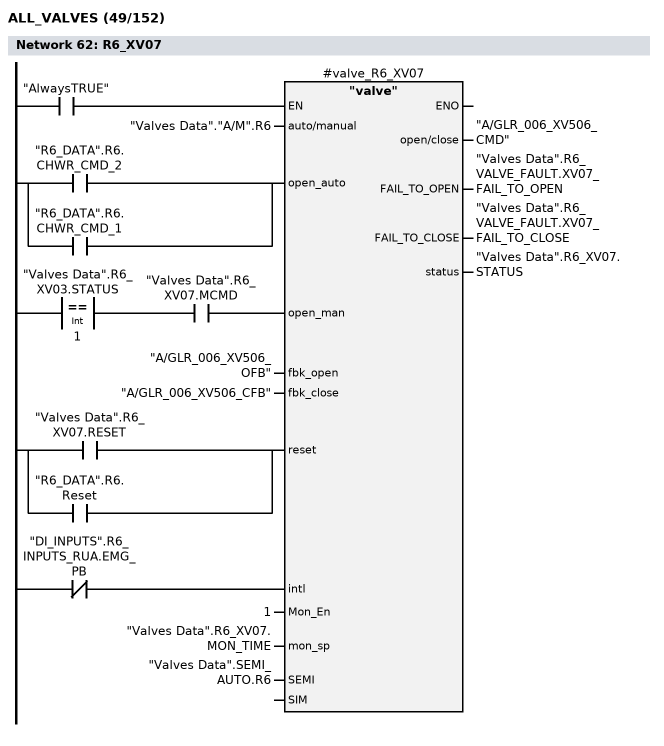
   RUNG wire#powerrail
      Contact( "AlwaysTRUE" )
      #valve_R6_XV07(open_auto := wire#w1, open_man := wire#w2, reset := wire#w3, intl := wire#w4, "auto/manual" := "Valves Data"."A/M".R6, fbk_open := "A/GLR_006_XV506_OFB", fbk_close := "A/GLR_006_XV506_CFB", Mon_En := 1, mon_sp := "Valves Data".R6_XV07.MON_TIME, SEMI := "Valves Data".SEMI_AUTO.R6, SIM :=, "open/close" => "A/GLR_006_XV506_CMD", FAIL_TO_OPEN => "Valves Data".R6_VALVE_FAULT.XV07_FAIL_TO_OPEN, FAIL_TO_CLOSE => "Valves Data".R6_VALVE_FAULT.XV07_FAIL_TO_CLOSE, status => "Valves Data".R6_XV07.STATUS)
   END_RUNG
   RUNG wire#powerrail
      Contact( "R6_DATA".R6.CHWR_CMD_2 )
   END_RUNG wire#w1
   RUNG wire#powerrail
      Contact( "R6_DATA".R6.CHWR_CMD_1 )
   END_RUNG wire#w1
   RUNG wire#powerrail
      { S7_Templates := "SrcType := Int" } EQ_Contact(in1 := "Valves Data".R6_XV03.STATUS, in2 := 1)
      Contact( "Valves Data".R6_XV07.MCMD )
   END_RUNG wire#w2
   RUNG wire#powerrail
      Contact( "Valves Data".R6_XV07.RESET )
   END_RUNG wire#w3
   RUNG wire#powerrail
      Contact( "R6_DATA".R6.Reset )
   END_RUNG wire#w3
   RUNG wire#powerrail
      I_Contact( "DI_INPUTS".R6_INPUTS_RUA.EMG_PB )
   END_RUNG wire#w4
   // the same network as SCL:
   IF "AlwaysTRUE" THEN
       #valve_R6_XV07("auto/manual" := "Valves Data"."A/M".R6,   // "valve"
                      open_auto := "R6_DATA".R6.CHWR_CMD_2 OR "R6_DATA".R6.CHWR_CMD_1,
                      open_man := ("Valves Data".R6_XV03.STATUS = 1) AND "Valves Data".R6_XV07.MCMD,
                      fbk_open := "A/GLR_006_XV506_OFB",
                      fbk_close := "A/GLR_006_XV506_CFB",
                      reset := "Valves Data".R6_XV07.RESET OR "R6_DATA".R6.Reset,
                      intl := NOT "DI_INPUTS".R6_INPUTS_RUA.EMG_PB,
                      Mon_En := 1,
                      mon_sp := "Valves Data".R6_XV07.MON_TIME,
                      SEMI := "Valves Data".SEMI_AUTO.R6,
                      "open/close" => "A/GLR_006_XV506_CMD",
                      FAIL_TO_OPEN => "Valves Data".R6_VALVE_FAULT.XV07_FAIL_TO_OPEN,
                      FAIL_TO_CLOSE => "Valves Data".R6_VALVE_FAULT.XV07_FAIL_TO_CLOSE,
                      status => "Valves Data".R6_XV07.STATUS);
   END_IF;
END_REGION

REGION Network 63: R6_XV08
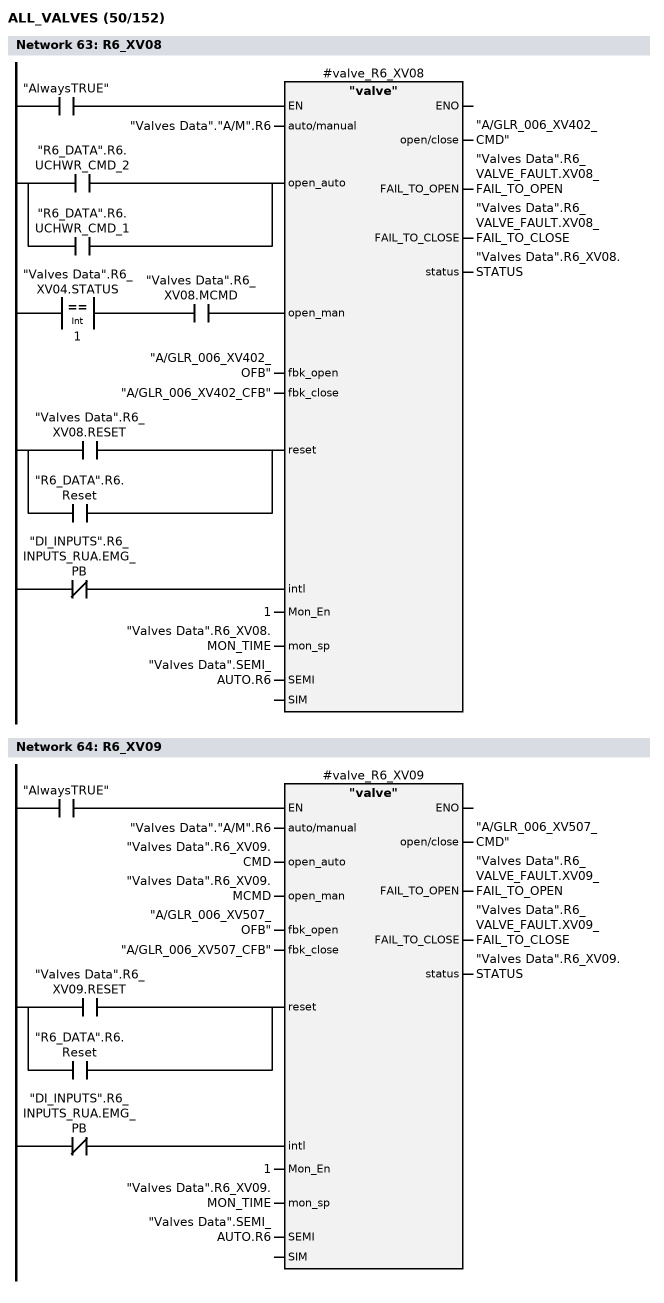
   RUNG wire#powerrail
      Contact( "AlwaysTRUE" )
      #valve_R6_XV08(open_auto := wire#w1, open_man := wire#w2, reset := wire#w3, intl := wire#w4, "auto/manual" := "Valves Data"."A/M".R6, fbk_open := "A/GLR_006_XV402_OFB", fbk_close := "A/GLR_006_XV402_CFB", Mon_En := 1, mon_sp := "Valves Data".R6_XV08.MON_TIME, SEMI := "Valves Data".SEMI_AUTO.R6, SIM :=, "open/close" => "A/GLR_006_XV402_CMD", FAIL_TO_OPEN => "Valves Data".R6_VALVE_FAULT.XV08_FAIL_TO_OPEN, FAIL_TO_CLOSE => "Valves Data".R6_VALVE_FAULT.XV08_FAIL_TO_CLOSE, status => "Valves Data".R6_XV08.STATUS)
   END_RUNG
   RUNG wire#powerrail
      Contact( "R6_DATA".R6.UCHWR_CMD_2 )
   END_RUNG wire#w1
   RUNG wire#powerrail
      Contact( "R6_DATA".R6.UCHWR_CMD_1 )
   END_RUNG wire#w1
   RUNG wire#powerrail
      { S7_Templates := "SrcType := Int" } EQ_Contact(in1 := "Valves Data".R6_XV04.STATUS, in2 := 1)
      Contact( "Valves Data".R6_XV08.MCMD )
   END_RUNG wire#w2
   RUNG wire#powerrail
      Contact( "Valves Data".R6_XV08.RESET )
   END_RUNG wire#w3
   RUNG wire#powerrail
      Contact( "R6_DATA".R6.Reset )
   END_RUNG wire#w3
   RUNG wire#powerrail
      I_Contact( "DI_INPUTS".R6_INPUTS_RUA.EMG_PB )
   END_RUNG wire#w4
   // the same network as SCL:
   IF "AlwaysTRUE" THEN
       #valve_R6_XV08("auto/manual" := "Valves Data"."A/M".R6,   // "valve"
                      open_auto := "R6_DATA".R6.UCHWR_CMD_2 OR "R6_DATA".R6.UCHWR_CMD_1,
                      open_man := ("Valves Data".R6_XV04.STATUS = 1) AND "Valves Data".R6_XV08.MCMD,
                      fbk_open := "A/GLR_006_XV402_OFB",
                      fbk_close := "A/GLR_006_XV402_CFB",
                      reset := "Valves Data".R6_XV08.RESET OR "R6_DATA".R6.Reset,
                      intl := NOT "DI_INPUTS".R6_INPUTS_RUA.EMG_PB,
                      Mon_En := 1,
                      mon_sp := "Valves Data".R6_XV08.MON_TIME,
                      SEMI := "Valves Data".SEMI_AUTO.R6,
                      "open/close" => "A/GLR_006_XV402_CMD",
                      FAIL_TO_OPEN => "Valves Data".R6_VALVE_FAULT.XV08_FAIL_TO_OPEN,
                      FAIL_TO_CLOSE => "Valves Data".R6_VALVE_FAULT.XV08_FAIL_TO_CLOSE,
                      status => "Valves Data".R6_XV08.STATUS);
   END_IF;
END_REGION

REGION Network 64: R6_XV09
   RUNG wire#powerrail
      Contact( "AlwaysTRUE" )
      #valve_R6_XV09(reset := wire#w1, intl := wire#w2, "auto/manual" := "Valves Data"."A/M".R6, open_auto := "Valves Data".R6_XV09.CMD, open_man := "Valves Data".R6_XV09.MCMD, fbk_open := "A/GLR_006_XV507_OFB", fbk_close := "A/GLR_006_XV507_CFB", Mon_En := 1, mon_sp := "Valves Data".R6_XV09.MON_TIME, SEMI := "Valves Data".SEMI_AUTO.R6, SIM :=, "open/close" => "A/GLR_006_XV507_CMD", FAIL_TO_OPEN => "Valves Data".R6_VALVE_FAULT.XV09_FAIL_TO_OPEN, FAIL_TO_CLOSE => "Valves Data".R6_VALVE_FAULT.XV09_FAIL_TO_CLOSE, status => "Valves Data".R6_XV09.STATUS)
   END_RUNG
   RUNG wire#powerrail
      Contact( "Valves Data".R6_XV09.RESET )
   END_RUNG wire#w1
   RUNG wire#powerrail
      Contact( "R6_DATA".R6.Reset )
   END_RUNG wire#w1
   RUNG wire#powerrail
      I_Contact( "DI_INPUTS".R6_INPUTS_RUA.EMG_PB )
   END_RUNG wire#w2
   // the same network as SCL:
   IF "AlwaysTRUE" THEN
       #valve_R6_XV09("auto/manual" := "Valves Data"."A/M".R6,   // "valve"
                      open_auto := "Valves Data".R6_XV09.CMD,
                      open_man := "Valves Data".R6_XV09.MCMD,
                      fbk_open := "A/GLR_006_XV507_OFB",
                      fbk_close := "A/GLR_006_XV507_CFB",
                      reset := "Valves Data".R6_XV09.RESET OR "R6_DATA".R6.Reset,
                      intl := NOT "DI_INPUTS".R6_INPUTS_RUA.EMG_PB,
                      Mon_En := 1,
                      mon_sp := "Valves Data".R6_XV09.MON_TIME,
                      SEMI := "Valves Data".SEMI_AUTO.R6,
                      "open/close" => "A/GLR_006_XV507_CMD",
                      FAIL_TO_OPEN => "Valves Data".R6_VALVE_FAULT.XV09_FAIL_TO_OPEN,
                      FAIL_TO_CLOSE => "Valves Data".R6_VALVE_FAULT.XV09_FAIL_TO_CLOSE,
                      status => "Valves Data".R6_XV09.STATUS);
   END_IF;
END_REGION

REGION Network 65: R6_XV10
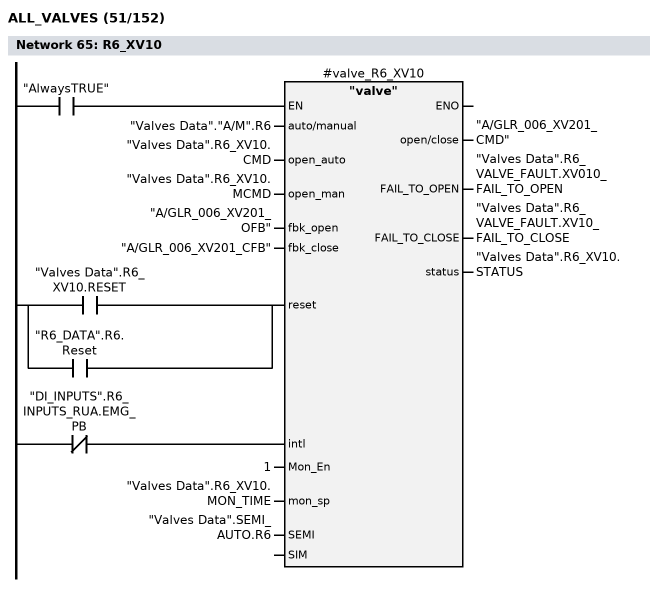
   RUNG wire#powerrail
      Contact( "AlwaysTRUE" )
      #valve_R6_XV10(reset := wire#w1, intl := wire#w2, "auto/manual" := "Valves Data"."A/M".R6, open_auto := "Valves Data".R6_XV10.CMD, open_man := "Valves Data".R6_XV10.MCMD, fbk_open := "A/GLR_006_XV201_OFB", fbk_close := "A/GLR_006_XV201_CFB", Mon_En := 1, mon_sp := "Valves Data".R6_XV10.MON_TIME, SEMI := "Valves Data".SEMI_AUTO.R6, SIM :=, "open/close" => "A/GLR_006_XV201_CMD", FAIL_TO_OPEN => "Valves Data".R6_VALVE_FAULT.XV010_FAIL_TO_OPEN, FAIL_TO_CLOSE => "Valves Data".R6_VALVE_FAULT.XV10_FAIL_TO_CLOSE, status => "Valves Data".R6_XV10.STATUS)
   END_RUNG
   RUNG wire#powerrail
      Contact( "Valves Data".R6_XV10.RESET )
   END_RUNG wire#w1
   RUNG wire#powerrail
      Contact( "R6_DATA".R6.Reset )
   END_RUNG wire#w1
   RUNG wire#powerrail
      I_Contact( "DI_INPUTS".R6_INPUTS_RUA.EMG_PB )
   END_RUNG wire#w2
   // the same network as SCL:
   IF "AlwaysTRUE" THEN
       #valve_R6_XV10("auto/manual" := "Valves Data"."A/M".R6,   // "valve"
                      open_auto := "Valves Data".R6_XV10.CMD,
                      open_man := "Valves Data".R6_XV10.MCMD,
                      fbk_open := "A/GLR_006_XV201_OFB",
                      fbk_close := "A/GLR_006_XV201_CFB",
                      reset := "Valves Data".R6_XV10.RESET OR "R6_DATA".R6.Reset,
                      intl := NOT "DI_INPUTS".R6_INPUTS_RUA.EMG_PB,
                      Mon_En := 1,
                      mon_sp := "Valves Data".R6_XV10.MON_TIME,
                      SEMI := "Valves Data".SEMI_AUTO.R6,
                      "open/close" => "A/GLR_006_XV201_CMD",
                      FAIL_TO_OPEN => "Valves Data".R6_VALVE_FAULT.XV010_FAIL_TO_OPEN,
                      FAIL_TO_CLOSE => "Valves Data".R6_VALVE_FAULT.XV10_FAIL_TO_CLOSE,
                      status => "Valves Data".R6_XV10.STATUS);
   END_IF;
END_REGION

REGION Network 66: ****REACTOR_07****
END_REGION

REGION Network 67: R7_XV01
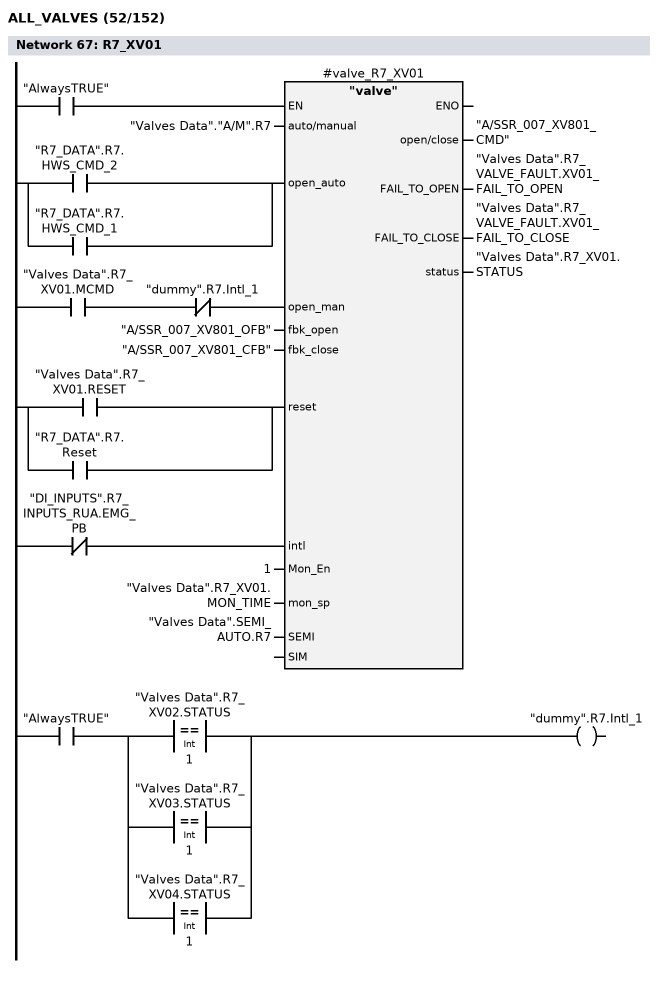
   RUNG wire#powerrail
      Contact( "AlwaysTRUE" )
      #valve_R7_XV01(open_auto := wire#w1, open_man := wire#w2, reset := wire#w3, intl := wire#w4, "auto/manual" := "Valves Data"."A/M".R7, fbk_open := "A/SSR_007_XV801_OFB", fbk_close := "A/SSR_007_XV801_CFB", Mon_En := 1, mon_sp := "Valves Data".R7_XV01.MON_TIME, SEMI := "Valves Data".SEMI_AUTO.R7, SIM :=, "open/close" => "A/SSR_007_XV801_CMD", FAIL_TO_OPEN => "Valves Data".R7_VALVE_FAULT.XV01_FAIL_TO_OPEN, FAIL_TO_CLOSE => "Valves Data".R7_VALVE_FAULT.XV01_FAIL_TO_CLOSE, status => "Valves Data".R7_XV01.STATUS)
   END_RUNG
   RUNG wire#powerrail
      Contact( "R7_DATA".R7.HWS_CMD_2 )
   END_RUNG wire#w1
   RUNG wire#powerrail
      Contact( "R7_DATA".R7.HWS_CMD_1 )
   END_RUNG wire#w1
   RUNG wire#powerrail
      Contact( "Valves Data".R7_XV01.MCMD )
      I_Contact( "dummy".R7.Intl_1 )
   END_RUNG wire#w2
   RUNG wire#powerrail
      Contact( "Valves Data".R7_XV01.RESET )
   END_RUNG wire#w3
   RUNG wire#powerrail
      Contact( "R7_DATA".R7.Reset )
   END_RUNG wire#w3
   RUNG wire#powerrail
      I_Contact( "DI_INPUTS".R7_INPUTS_RUA.EMG_PB )
   END_RUNG wire#w4
   RUNG wire#powerrail
      Contact( "AlwaysTRUE" )
      wire#w5
      { S7_Templates := "SrcType := Int" } EQ_Contact(in1 := "Valves Data".R7_XV02.STATUS, in2 := 1)
      wire#w6
      Coil( "dummy".R7.Intl_1 )
   END_RUNG
   RUNG wire#w5
      { S7_Templates := "SrcType := Int" } EQ_Contact(in1 := "Valves Data".R7_XV03.STATUS, in2 := 1)
   END_RUNG wire#w6
   RUNG wire#w5
      { S7_Templates := "SrcType := Int" } EQ_Contact(in1 := "Valves Data".R7_XV04.STATUS, in2 := 1)
   END_RUNG wire#w6
   // the same network as SCL:
   IF "AlwaysTRUE" THEN
       #valve_R7_XV01("auto/manual" := "Valves Data"."A/M".R7,   // "valve"
                      open_auto := "R7_DATA".R7.HWS_CMD_2 OR "R7_DATA".R7.HWS_CMD_1,
                      open_man := "Valves Data".R7_XV01.MCMD AND NOT "dummy".R7.Intl_1,
                      fbk_open := "A/SSR_007_XV801_OFB",
                      fbk_close := "A/SSR_007_XV801_CFB",
                      reset := "Valves Data".R7_XV01.RESET OR "R7_DATA".R7.Reset,
                      intl := NOT "DI_INPUTS".R7_INPUTS_RUA.EMG_PB,
                      Mon_En := 1,
                      mon_sp := "Valves Data".R7_XV01.MON_TIME,
                      SEMI := "Valves Data".SEMI_AUTO.R7,
                      "open/close" => "A/SSR_007_XV801_CMD",
                      FAIL_TO_OPEN => "Valves Data".R7_VALVE_FAULT.XV01_FAIL_TO_OPEN,
                      FAIL_TO_CLOSE => "Valves Data".R7_VALVE_FAULT.XV01_FAIL_TO_CLOSE,
                      status => "Valves Data".R7_XV01.STATUS);
   END_IF;
   "dummy".R7.Intl_1 := "AlwaysTRUE" AND (("Valves Data".R7_XV02.STATUS = 1) OR ("Valves Data".R7_XV03.STATUS = 1) OR ("Valves Data".R7_XV04.STATUS = 1));
END_REGION

REGION Network 68: R7_XV02
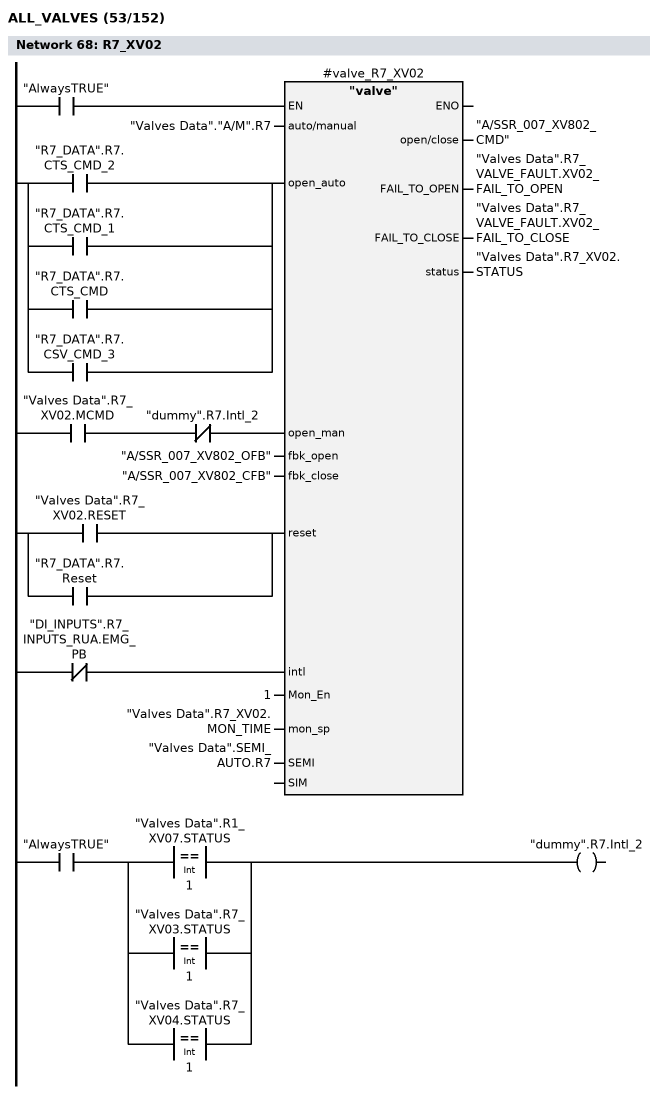
   RUNG wire#powerrail
      Contact( "AlwaysTRUE" )
      #valve_R7_XV02(open_auto := wire#w1, open_man := wire#w2, reset := wire#w3, intl := wire#w4, "auto/manual" := "Valves Data"."A/M".R7, fbk_open := "A/SSR_007_XV802_OFB", fbk_close := "A/SSR_007_XV802_CFB", Mon_En := 1, mon_sp := "Valves Data".R7_XV02.MON_TIME, SEMI := "Valves Data".SEMI_AUTO.R7, SIM :=, "open/close" => "A/SSR_007_XV802_CMD", FAIL_TO_OPEN => "Valves Data".R7_VALVE_FAULT.XV02_FAIL_TO_OPEN, FAIL_TO_CLOSE => "Valves Data".R7_VALVE_FAULT.XV02_FAIL_TO_CLOSE, status => "Valves Data".R7_XV02.STATUS)
   END_RUNG
   RUNG wire#powerrail
      Contact( "R7_DATA".R7.CTS_CMD_2 )
   END_RUNG wire#w1
   RUNG wire#powerrail
      Contact( "R7_DATA".R7.CTS_CMD_1 )
   END_RUNG wire#w1
   RUNG wire#powerrail
      Contact( "R7_DATA".R7.CTS_CMD )
   END_RUNG wire#w1
   RUNG wire#powerrail
      Contact( "R7_DATA".R7.CSV_CMD_3 )
   END_RUNG wire#w1
   RUNG wire#powerrail
      Contact( "Valves Data".R7_XV02.MCMD )
      I_Contact( "dummy".R7.Intl_2 )
   END_RUNG wire#w2
   RUNG wire#powerrail
      Contact( "Valves Data".R7_XV02.RESET )
   END_RUNG wire#w3
   RUNG wire#powerrail
      Contact( "R7_DATA".R7.Reset )
   END_RUNG wire#w3
   RUNG wire#powerrail
      I_Contact( "DI_INPUTS".R7_INPUTS_RUA.EMG_PB )
   END_RUNG wire#w4
   RUNG wire#powerrail
      Contact( "AlwaysTRUE" )
      wire#w5
      { S7_Templates := "SrcType := Int" } EQ_Contact(in1 := "Valves Data".R1_XV07.STATUS, in2 := 1)
      wire#w6
      Coil( "dummy".R7.Intl_2 )
   END_RUNG
   RUNG wire#w5
      { S7_Templates := "SrcType := Int" } EQ_Contact(in1 := "Valves Data".R7_XV03.STATUS, in2 := 1)
   END_RUNG wire#w6
   RUNG wire#w5
      { S7_Templates := "SrcType := Int" } EQ_Contact(in1 := "Valves Data".R7_XV04.STATUS, in2 := 1)
   END_RUNG wire#w6
   // the same network as SCL:
   IF "AlwaysTRUE" THEN
       #valve_R7_XV02("auto/manual" := "Valves Data"."A/M".R7,   // "valve"
                      open_auto := "R7_DATA".R7.CTS_CMD_2 OR "R7_DATA".R7.CTS_CMD_1 OR "R7_DATA".R7.CTS_CMD OR "R7_DATA".R7.CSV_CMD_3,
                      open_man := "Valves Data".R7_XV02.MCMD AND NOT "dummy".R7.Intl_2,
                      fbk_open := "A/SSR_007_XV802_OFB",
                      fbk_close := "A/SSR_007_XV802_CFB",
                      reset := "Valves Data".R7_XV02.RESET OR "R7_DATA".R7.Reset,
                      intl := NOT "DI_INPUTS".R7_INPUTS_RUA.EMG_PB,
                      Mon_En := 1,
                      mon_sp := "Valves Data".R7_XV02.MON_TIME,
                      SEMI := "Valves Data".SEMI_AUTO.R7,
                      "open/close" => "A/SSR_007_XV802_CMD",
                      FAIL_TO_OPEN => "Valves Data".R7_VALVE_FAULT.XV02_FAIL_TO_OPEN,
                      FAIL_TO_CLOSE => "Valves Data".R7_VALVE_FAULT.XV02_FAIL_TO_CLOSE,
                      status => "Valves Data".R7_XV02.STATUS);
   END_IF;
   "dummy".R7.Intl_2 := "AlwaysTRUE" AND (("Valves Data".R1_XV07.STATUS = 1) OR ("Valves Data".R7_XV03.STATUS = 1) OR ("Valves Data".R7_XV04.STATUS = 1));
END_REGION

REGION Network 69: R7_XV03
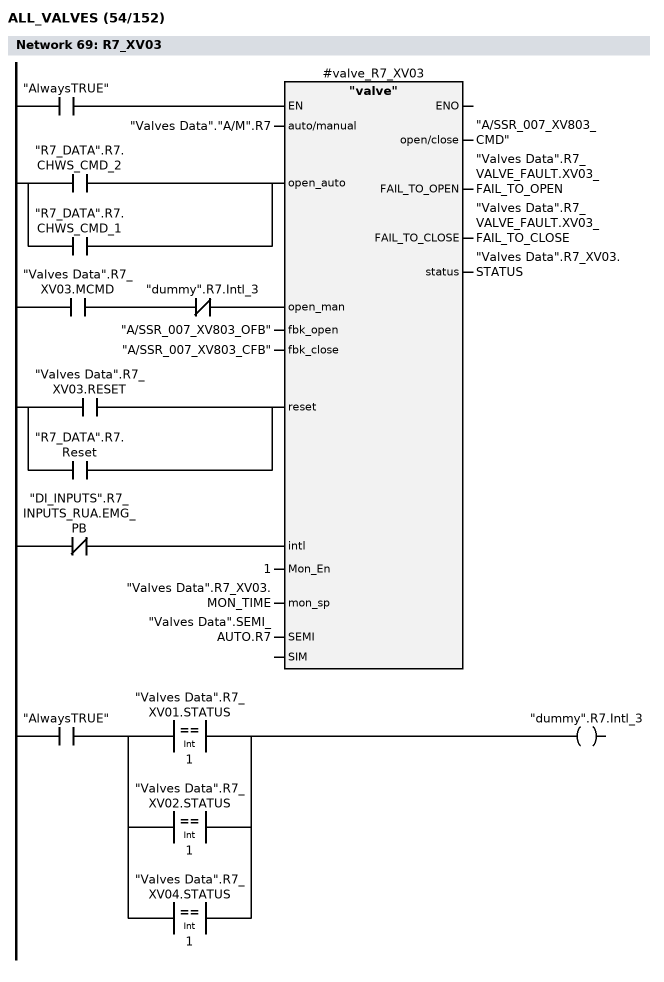
   RUNG wire#powerrail
      Contact( "AlwaysTRUE" )
      #valve_R7_XV03(open_auto := wire#w1, open_man := wire#w2, reset := wire#w3, intl := wire#w4, "auto/manual" := "Valves Data"."A/M".R7, fbk_open := "A/SSR_007_XV803_OFB", fbk_close := "A/SSR_007_XV803_CFB", Mon_En := 1, mon_sp := "Valves Data".R7_XV03.MON_TIME, SEMI := "Valves Data".SEMI_AUTO.R7, SIM :=, "open/close" => "A/SSR_007_XV803_CMD", FAIL_TO_OPEN => "Valves Data".R7_VALVE_FAULT.XV03_FAIL_TO_OPEN, FAIL_TO_CLOSE => "Valves Data".R7_VALVE_FAULT.XV03_FAIL_TO_CLOSE, status => "Valves Data".R7_XV03.STATUS)
   END_RUNG
   RUNG wire#powerrail
      Contact( "R7_DATA".R7.CHWS_CMD_2 )
   END_RUNG wire#w1
   RUNG wire#powerrail
      Contact( "R7_DATA".R7.CHWS_CMD_1 )
   END_RUNG wire#w1
   RUNG wire#powerrail
      Contact( "Valves Data".R7_XV03.MCMD )
      I_Contact( "dummy".R7.Intl_3 )
   END_RUNG wire#w2
   RUNG wire#powerrail
      Contact( "Valves Data".R7_XV03.RESET )
   END_RUNG wire#w3
   RUNG wire#powerrail
      Contact( "R7_DATA".R7.Reset )
   END_RUNG wire#w3
   RUNG wire#powerrail
      I_Contact( "DI_INPUTS".R7_INPUTS_RUA.EMG_PB )
   END_RUNG wire#w4
   RUNG wire#powerrail
      Contact( "AlwaysTRUE" )
      wire#w5
      { S7_Templates := "SrcType := Int" } EQ_Contact(in1 := "Valves Data".R7_XV01.STATUS, in2 := 1)
      wire#w6
      Coil( "dummy".R7.Intl_3 )
   END_RUNG
   RUNG wire#w5
      { S7_Templates := "SrcType := Int" } EQ_Contact(in1 := "Valves Data".R7_XV02.STATUS, in2 := 1)
   END_RUNG wire#w6
   RUNG wire#w5
      { S7_Templates := "SrcType := Int" } EQ_Contact(in1 := "Valves Data".R7_XV04.STATUS, in2 := 1)
   END_RUNG wire#w6
   // the same network as SCL:
   IF "AlwaysTRUE" THEN
       #valve_R7_XV03("auto/manual" := "Valves Data"."A/M".R7,   // "valve"
                      open_auto := "R7_DATA".R7.CHWS_CMD_2 OR "R7_DATA".R7.CHWS_CMD_1,
                      open_man := "Valves Data".R7_XV03.MCMD AND NOT "dummy".R7.Intl_3,
                      fbk_open := "A/SSR_007_XV803_OFB",
                      fbk_close := "A/SSR_007_XV803_CFB",
                      reset := "Valves Data".R7_XV03.RESET OR "R7_DATA".R7.Reset,
                      intl := NOT "DI_INPUTS".R7_INPUTS_RUA.EMG_PB,
                      Mon_En := 1,
                      mon_sp := "Valves Data".R7_XV03.MON_TIME,
                      SEMI := "Valves Data".SEMI_AUTO.R7,
                      "open/close" => "A/SSR_007_XV803_CMD",
                      FAIL_TO_OPEN => "Valves Data".R7_VALVE_FAULT.XV03_FAIL_TO_OPEN,
                      FAIL_TO_CLOSE => "Valves Data".R7_VALVE_FAULT.XV03_FAIL_TO_CLOSE,
                      status => "Valves Data".R7_XV03.STATUS);
   END_IF;
   "dummy".R7.Intl_3 := "AlwaysTRUE" AND (("Valves Data".R7_XV01.STATUS = 1) OR ("Valves Data".R7_XV02.STATUS = 1) OR ("Valves Data".R7_XV04.STATUS = 1));
END_REGION

REGION Network 70: R7_XV04
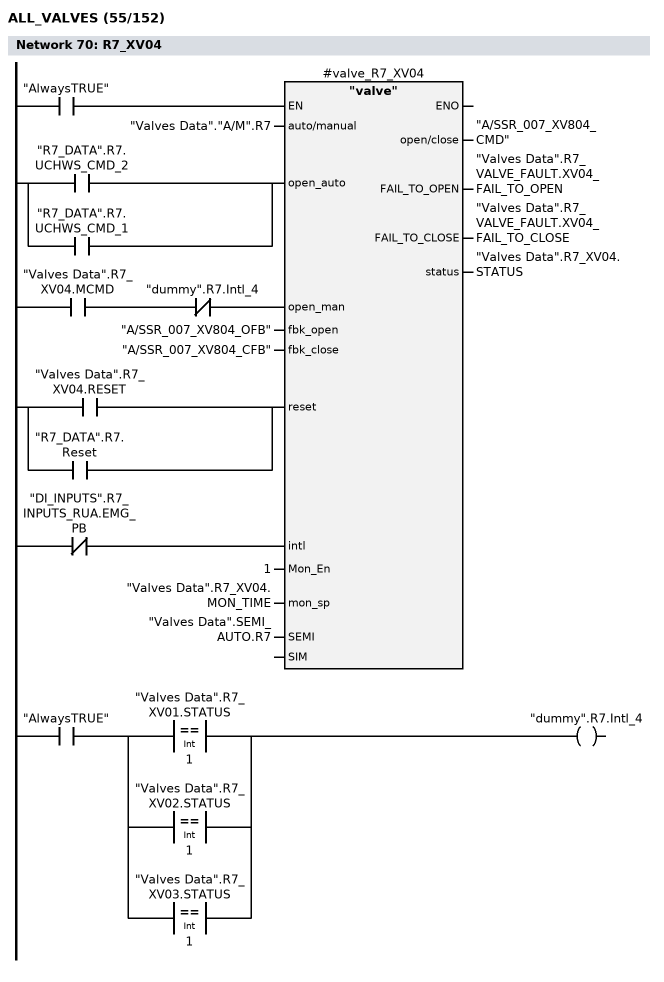
   RUNG wire#powerrail
      Contact( "AlwaysTRUE" )
      #valve_R7_XV04(open_auto := wire#w1, open_man := wire#w2, reset := wire#w3, intl := wire#w4, "auto/manual" := "Valves Data"."A/M".R7, fbk_open := "A/SSR_007_XV804_OFB", fbk_close := "A/SSR_007_XV804_CFB", Mon_En := 1, mon_sp := "Valves Data".R7_XV04.MON_TIME, SEMI := "Valves Data".SEMI_AUTO.R7, SIM :=, "open/close" => "A/SSR_007_XV804_CMD", FAIL_TO_OPEN => "Valves Data".R7_VALVE_FAULT.XV04_FAIL_TO_OPEN, FAIL_TO_CLOSE => "Valves Data".R7_VALVE_FAULT.XV04_FAIL_TO_CLOSE, status => "Valves Data".R7_XV04.STATUS)
   END_RUNG
   RUNG wire#powerrail
      Contact( "R7_DATA".R7.UCHWS_CMD_2 )
   END_RUNG wire#w1
   RUNG wire#powerrail
      Contact( "R7_DATA".R7.UCHWS_CMD_1 )
   END_RUNG wire#w1
   RUNG wire#powerrail
      Contact( "Valves Data".R7_XV04.MCMD )
      I_Contact( "dummy".R7.Intl_4 )
   END_RUNG wire#w2
   RUNG wire#powerrail
      Contact( "Valves Data".R7_XV04.RESET )
   END_RUNG wire#w3
   RUNG wire#powerrail
      Contact( "R7_DATA".R7.Reset )
   END_RUNG wire#w3
   RUNG wire#powerrail
      I_Contact( "DI_INPUTS".R7_INPUTS_RUA.EMG_PB )
   END_RUNG wire#w4
   RUNG wire#powerrail
      Contact( "AlwaysTRUE" )
      wire#w5
      { S7_Templates := "SrcType := Int" } EQ_Contact(in1 := "Valves Data".R7_XV01.STATUS, in2 := 1)
      wire#w6
      Coil( "dummy".R7.Intl_4 )
   END_RUNG
   RUNG wire#w5
      { S7_Templates := "SrcType := Int" } EQ_Contact(in1 := "Valves Data".R7_XV02.STATUS, in2 := 1)
   END_RUNG wire#w6
   RUNG wire#w5
      { S7_Templates := "SrcType := Int" } EQ_Contact(in1 := "Valves Data".R7_XV03.STATUS, in2 := 1)
   END_RUNG wire#w6
   // the same network as SCL:
   IF "AlwaysTRUE" THEN
       #valve_R7_XV04("auto/manual" := "Valves Data"."A/M".R7,   // "valve"
                      open_auto := "R7_DATA".R7.UCHWS_CMD_2 OR "R7_DATA".R7.UCHWS_CMD_1,
                      open_man := "Valves Data".R7_XV04.MCMD AND NOT "dummy".R7.Intl_4,
                      fbk_open := "A/SSR_007_XV804_OFB",
                      fbk_close := "A/SSR_007_XV804_CFB",
                      reset := "Valves Data".R7_XV04.RESET OR "R7_DATA".R7.Reset,
                      intl := NOT "DI_INPUTS".R7_INPUTS_RUA.EMG_PB,
                      Mon_En := 1,
                      mon_sp := "Valves Data".R7_XV04.MON_TIME,
                      SEMI := "Valves Data".SEMI_AUTO.R7,
                      "open/close" => "A/SSR_007_XV804_CMD",
                      FAIL_TO_OPEN => "Valves Data".R7_VALVE_FAULT.XV04_FAIL_TO_OPEN,
                      FAIL_TO_CLOSE => "Valves Data".R7_VALVE_FAULT.XV04_FAIL_TO_CLOSE,
                      status => "Valves Data".R7_XV04.STATUS);
   END_IF;
   "dummy".R7.Intl_4 := "AlwaysTRUE" AND (("Valves Data".R7_XV01.STATUS = 1) OR ("Valves Data".R7_XV02.STATUS = 1) OR ("Valves Data".R7_XV03.STATUS = 1));
END_REGION

REGION Network 71: R7_XV05
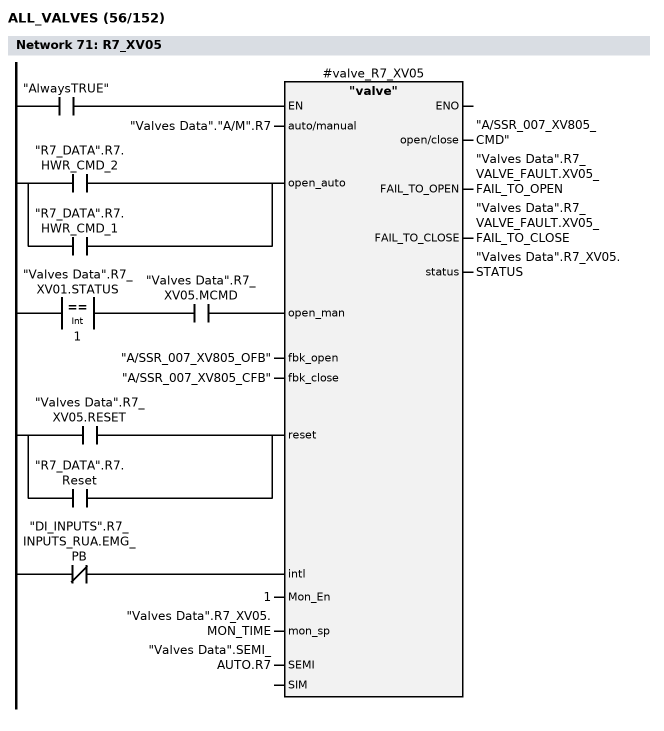
   RUNG wire#powerrail
      Contact( "AlwaysTRUE" )
      #valve_R7_XV05(open_auto := wire#w1, open_man := wire#w2, reset := wire#w3, intl := wire#w4, "auto/manual" := "Valves Data"."A/M".R7, fbk_open := "A/SSR_007_XV805_OFB", fbk_close := "A/SSR_007_XV805_CFB", Mon_En := 1, mon_sp := "Valves Data".R7_XV05.MON_TIME, SEMI := "Valves Data".SEMI_AUTO.R7, SIM :=, "open/close" => "A/SSR_007_XV805_CMD", FAIL_TO_OPEN => "Valves Data".R7_VALVE_FAULT.XV05_FAIL_TO_OPEN, FAIL_TO_CLOSE => "Valves Data".R7_VALVE_FAULT.XV05_FAIL_TO_CLOSE, status => "Valves Data".R7_XV05.STATUS)
   END_RUNG
   RUNG wire#powerrail
      Contact( "R7_DATA".R7.HWR_CMD_2 )
   END_RUNG wire#w1
   RUNG wire#powerrail
      Contact( "R7_DATA".R7.HWR_CMD_1 )
   END_RUNG wire#w1
   RUNG wire#powerrail
      { S7_Templates := "SrcType := Int" } EQ_Contact(in1 := "Valves Data".R7_XV01.STATUS, in2 := 1)
      Contact( "Valves Data".R7_XV05.MCMD )
   END_RUNG wire#w2
   RUNG wire#powerrail
      Contact( "Valves Data".R7_XV05.RESET )
   END_RUNG wire#w3
   RUNG wire#powerrail
      Contact( "R7_DATA".R7.Reset )
   END_RUNG wire#w3
   RUNG wire#powerrail
      I_Contact( "DI_INPUTS".R7_INPUTS_RUA.EMG_PB )
   END_RUNG wire#w4
   // the same network as SCL:
   IF "AlwaysTRUE" THEN
       #valve_R7_XV05("auto/manual" := "Valves Data"."A/M".R7,   // "valve"
                      open_auto := "R7_DATA".R7.HWR_CMD_2 OR "R7_DATA".R7.HWR_CMD_1,
                      open_man := ("Valves Data".R7_XV01.STATUS = 1) AND "Valves Data".R7_XV05.MCMD,
                      fbk_open := "A/SSR_007_XV805_OFB",
                      fbk_close := "A/SSR_007_XV805_CFB",
                      reset := "Valves Data".R7_XV05.RESET OR "R7_DATA".R7.Reset,
                      intl := NOT "DI_INPUTS".R7_INPUTS_RUA.EMG_PB,
                      Mon_En := 1,
                      mon_sp := "Valves Data".R7_XV05.MON_TIME,
                      SEMI := "Valves Data".SEMI_AUTO.R7,
                      "open/close" => "A/SSR_007_XV805_CMD",
                      FAIL_TO_OPEN => "Valves Data".R7_VALVE_FAULT.XV05_FAIL_TO_OPEN,
                      FAIL_TO_CLOSE => "Valves Data".R7_VALVE_FAULT.XV05_FAIL_TO_CLOSE,
                      status => "Valves Data".R7_XV05.STATUS);
   END_IF;
END_REGION

REGION Network 72: R7_XV06
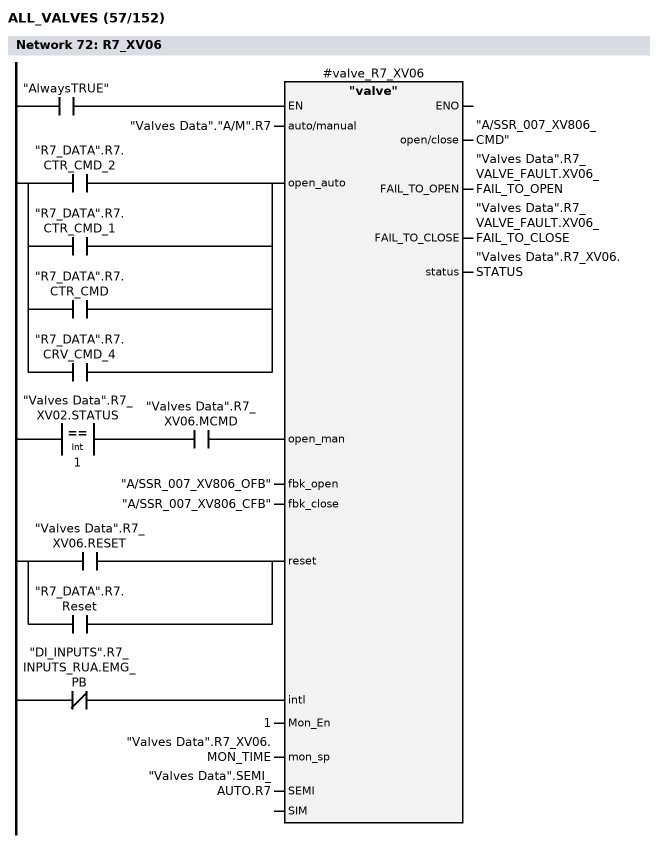
   RUNG wire#powerrail
      Contact( "AlwaysTRUE" )
      #valve_R7_XV06(open_auto := wire#w1, open_man := wire#w2, reset := wire#w3, intl := wire#w4, "auto/manual" := "Valves Data"."A/M".R7, fbk_open := "A/SSR_007_XV806_OFB", fbk_close := "A/SSR_007_XV806_CFB", Mon_En := 1, mon_sp := "Valves Data".R7_XV06.MON_TIME, SEMI := "Valves Data".SEMI_AUTO.R7, SIM :=, "open/close" => "A/SSR_007_XV806_CMD", FAIL_TO_OPEN => "Valves Data".R7_VALVE_FAULT.XV06_FAIL_TO_OPEN, FAIL_TO_CLOSE => "Valves Data".R7_VALVE_FAULT.XV06_FAIL_TO_CLOSE, status => "Valves Data".R7_XV06.STATUS)
   END_RUNG
   RUNG wire#powerrail
      Contact( "R7_DATA".R7.CTR_CMD_2 )
   END_RUNG wire#w1
   RUNG wire#powerrail
      Contact( "R7_DATA".R7.CTR_CMD_1 )
   END_RUNG wire#w1
   RUNG wire#powerrail
      Contact( "R7_DATA".R7.CTR_CMD )
   END_RUNG wire#w1
   RUNG wire#powerrail
      Contact( "R7_DATA".R7.CRV_CMD_4 )
   END_RUNG wire#w1
   RUNG wire#powerrail
      { S7_Templates := "SrcType := Int" } EQ_Contact(in1 := "Valves Data".R7_XV02.STATUS, in2 := 1)
      Contact( "Valves Data".R7_XV06.MCMD )
   END_RUNG wire#w2
   RUNG wire#powerrail
      Contact( "Valves Data".R7_XV06.RESET )
   END_RUNG wire#w3
   RUNG wire#powerrail
      Contact( "R7_DATA".R7.Reset )
   END_RUNG wire#w3
   RUNG wire#powerrail
      I_Contact( "DI_INPUTS".R7_INPUTS_RUA.EMG_PB )
   END_RUNG wire#w4
   // the same network as SCL:
   IF "AlwaysTRUE" THEN
       #valve_R7_XV06("auto/manual" := "Valves Data"."A/M".R7,   // "valve"
                      open_auto := "R7_DATA".R7.CTR_CMD_2 OR "R7_DATA".R7.CTR_CMD_1 OR "R7_DATA".R7.CTR_CMD OR "R7_DATA".R7.CRV_CMD_4,
                      open_man := ("Valves Data".R7_XV02.STATUS = 1) AND "Valves Data".R7_XV06.MCMD,
                      fbk_open := "A/SSR_007_XV806_OFB",
                      fbk_close := "A/SSR_007_XV806_CFB",
                      reset := "Valves Data".R7_XV06.RESET OR "R7_DATA".R7.Reset,
                      intl := NOT "DI_INPUTS".R7_INPUTS_RUA.EMG_PB,
                      Mon_En := 1,
                      mon_sp := "Valves Data".R7_XV06.MON_TIME,
                      SEMI := "Valves Data".SEMI_AUTO.R7,
                      "open/close" => "A/SSR_007_XV806_CMD",
                      FAIL_TO_OPEN => "Valves Data".R7_VALVE_FAULT.XV06_FAIL_TO_OPEN,
                      FAIL_TO_CLOSE => "Valves Data".R7_VALVE_FAULT.XV06_FAIL_TO_CLOSE,
                      status => "Valves Data".R7_XV06.STATUS);
   END_IF;
END_REGION

REGION Network 73: R7_XV07
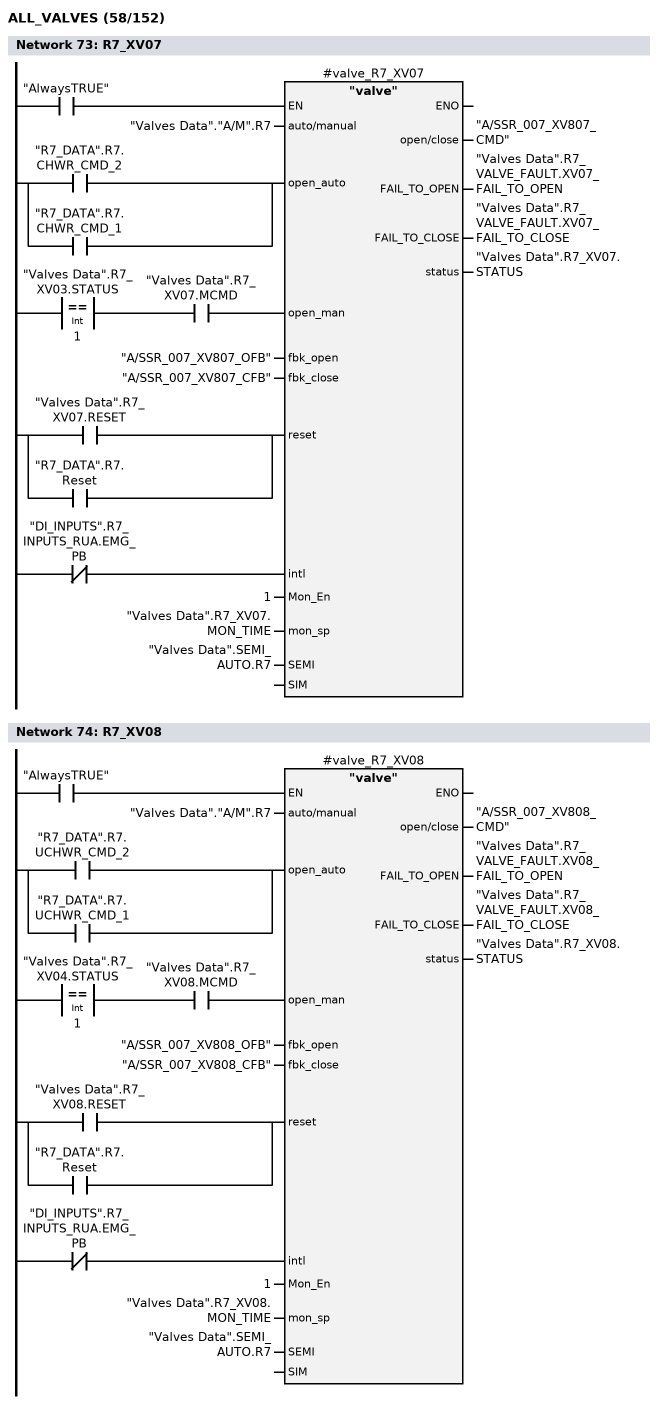
   RUNG wire#powerrail
      Contact( "AlwaysTRUE" )
      #valve_R7_XV07(open_auto := wire#w1, open_man := wire#w2, reset := wire#w3, intl := wire#w4, "auto/manual" := "Valves Data"."A/M".R7, fbk_open := "A/SSR_007_XV807_OFB", fbk_close := "A/SSR_007_XV807_CFB", Mon_En := 1, mon_sp := "Valves Data".R7_XV07.MON_TIME, SEMI := "Valves Data".SEMI_AUTO.R7, SIM :=, "open/close" => "A/SSR_007_XV807_CMD", FAIL_TO_OPEN => "Valves Data".R7_VALVE_FAULT.XV07_FAIL_TO_OPEN, FAIL_TO_CLOSE => "Valves Data".R7_VALVE_FAULT.XV07_FAIL_TO_CLOSE, status => "Valves Data".R7_XV07.STATUS)
   END_RUNG
   RUNG wire#powerrail
      Contact( "R7_DATA".R7.CHWR_CMD_2 )
   END_RUNG wire#w1
   RUNG wire#powerrail
      Contact( "R7_DATA".R7.CHWR_CMD_1 )
   END_RUNG wire#w1
   RUNG wire#powerrail
      { S7_Templates := "SrcType := Int" } EQ_Contact(in1 := "Valves Data".R7_XV03.STATUS, in2 := 1)
      Contact( "Valves Data".R7_XV07.MCMD )
   END_RUNG wire#w2
   RUNG wire#powerrail
      Contact( "Valves Data".R7_XV07.RESET )
   END_RUNG wire#w3
   RUNG wire#powerrail
      Contact( "R7_DATA".R7.Reset )
   END_RUNG wire#w3
   RUNG wire#powerrail
      I_Contact( "DI_INPUTS".R7_INPUTS_RUA.EMG_PB )
   END_RUNG wire#w4
   // the same network as SCL:
   IF "AlwaysTRUE" THEN
       #valve_R7_XV07("auto/manual" := "Valves Data"."A/M".R7,   // "valve"
                      open_auto := "R7_DATA".R7.CHWR_CMD_2 OR "R7_DATA".R7.CHWR_CMD_1,
                      open_man := ("Valves Data".R7_XV03.STATUS = 1) AND "Valves Data".R7_XV07.MCMD,
                      fbk_open := "A/SSR_007_XV807_OFB",
                      fbk_close := "A/SSR_007_XV807_CFB",
                      reset := "Valves Data".R7_XV07.RESET OR "R7_DATA".R7.Reset,
                      intl := NOT "DI_INPUTS".R7_INPUTS_RUA.EMG_PB,
                      Mon_En := 1,
                      mon_sp := "Valves Data".R7_XV07.MON_TIME,
                      SEMI := "Valves Data".SEMI_AUTO.R7,
                      "open/close" => "A/SSR_007_XV807_CMD",
                      FAIL_TO_OPEN => "Valves Data".R7_VALVE_FAULT.XV07_FAIL_TO_OPEN,
                      FAIL_TO_CLOSE => "Valves Data".R7_VALVE_FAULT.XV07_FAIL_TO_CLOSE,
                      status => "Valves Data".R7_XV07.STATUS);
   END_IF;
END_REGION

REGION Network 74: R7_XV08
   RUNG wire#powerrail
      Contact( "AlwaysTRUE" )
      #valve_R7_XV08(open_auto := wire#w1, open_man := wire#w2, reset := wire#w3, intl := wire#w4, "auto/manual" := "Valves Data"."A/M".R7, fbk_open := "A/SSR_007_XV808_OFB", fbk_close := "A/SSR_007_XV808_CFB", Mon_En := 1, mon_sp := "Valves Data".R7_XV08.MON_TIME, SEMI := "Valves Data".SEMI_AUTO.R7, SIM :=, "open/close" => "A/SSR_007_XV808_CMD", FAIL_TO_OPEN => "Valves Data".R7_VALVE_FAULT.XV08_FAIL_TO_OPEN, FAIL_TO_CLOSE => "Valves Data".R7_VALVE_FAULT.XV08_FAIL_TO_CLOSE, status => "Valves Data".R7_XV08.STATUS)
   END_RUNG
   RUNG wire#powerrail
      Contact( "R7_DATA".R7.UCHWR_CMD_2 )
   END_RUNG wire#w1
   RUNG wire#powerrail
      Contact( "R7_DATA".R7.UCHWR_CMD_1 )
   END_RUNG wire#w1
   RUNG wire#powerrail
      { S7_Templates := "SrcType := Int" } EQ_Contact(in1 := "Valves Data".R7_XV04.STATUS, in2 := 1)
      Contact( "Valves Data".R7_XV08.MCMD )
   END_RUNG wire#w2
   RUNG wire#powerrail
      Contact( "Valves Data".R7_XV08.RESET )
   END_RUNG wire#w3
   RUNG wire#powerrail
      Contact( "R7_DATA".R7.Reset )
   END_RUNG wire#w3
   RUNG wire#powerrail
      I_Contact( "DI_INPUTS".R7_INPUTS_RUA.EMG_PB )
   END_RUNG wire#w4
   // the same network as SCL:
   IF "AlwaysTRUE" THEN
       #valve_R7_XV08("auto/manual" := "Valves Data"."A/M".R7,   // "valve"
                      open_auto := "R7_DATA".R7.UCHWR_CMD_2 OR "R7_DATA".R7.UCHWR_CMD_1,
                      open_man := ("Valves Data".R7_XV04.STATUS = 1) AND "Valves Data".R7_XV08.MCMD,
                      fbk_open := "A/SSR_007_XV808_OFB",
                      fbk_close := "A/SSR_007_XV808_CFB",
                      reset := "Valves Data".R7_XV08.RESET OR "R7_DATA".R7.Reset,
                      intl := NOT "DI_INPUTS".R7_INPUTS_RUA.EMG_PB,
                      Mon_En := 1,
                      mon_sp := "Valves Data".R7_XV08.MON_TIME,
                      SEMI := "Valves Data".SEMI_AUTO.R7,
                      "open/close" => "A/SSR_007_XV808_CMD",
                      FAIL_TO_OPEN => "Valves Data".R7_VALVE_FAULT.XV08_FAIL_TO_OPEN,
                      FAIL_TO_CLOSE => "Valves Data".R7_VALVE_FAULT.XV08_FAIL_TO_CLOSE,
                      status => "Valves Data".R7_XV08.STATUS);
   END_IF;
END_REGION

REGION Network 75: R7_XV09
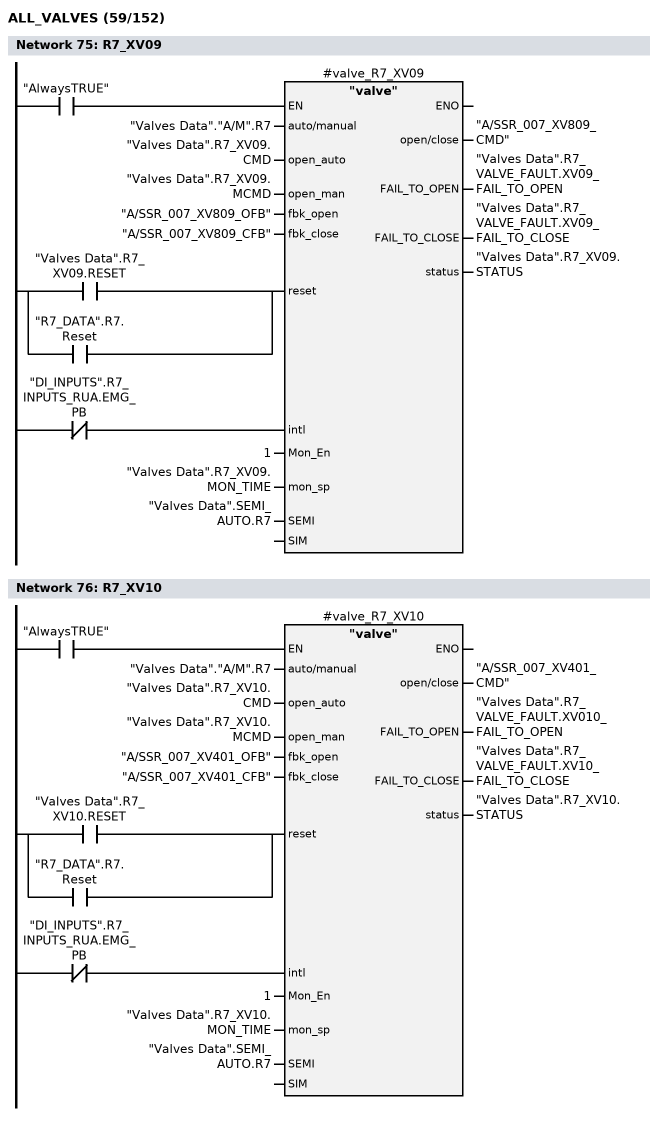
   RUNG wire#powerrail
      Contact( "AlwaysTRUE" )
      #valve_R7_XV09(reset := wire#w1, intl := wire#w2, "auto/manual" := "Valves Data"."A/M".R7, open_auto := "Valves Data".R7_XV09.CMD, open_man := "Valves Data".R7_XV09.MCMD, fbk_open := "A/SSR_007_XV809_OFB", fbk_close := "A/SSR_007_XV809_CFB", Mon_En := 1, mon_sp := "Valves Data".R7_XV09.MON_TIME, SEMI := "Valves Data".SEMI_AUTO.R7, SIM :=, "open/close" => "A/SSR_007_XV809_CMD", FAIL_TO_OPEN => "Valves Data".R7_VALVE_FAULT.XV09_FAIL_TO_OPEN, FAIL_TO_CLOSE => "Valves Data".R7_VALVE_FAULT.XV09_FAIL_TO_CLOSE, status => "Valves Data".R7_XV09.STATUS)
   END_RUNG
   RUNG wire#powerrail
      Contact( "Valves Data".R7_XV09.RESET )
   END_RUNG wire#w1
   RUNG wire#powerrail
      Contact( "R7_DATA".R7.Reset )
   END_RUNG wire#w1
   RUNG wire#powerrail
      I_Contact( "DI_INPUTS".R7_INPUTS_RUA.EMG_PB )
   END_RUNG wire#w2
   // the same network as SCL:
   IF "AlwaysTRUE" THEN
       #valve_R7_XV09("auto/manual" := "Valves Data"."A/M".R7,   // "valve"
                      open_auto := "Valves Data".R7_XV09.CMD,
                      open_man := "Valves Data".R7_XV09.MCMD,
                      fbk_open := "A/SSR_007_XV809_OFB",
                      fbk_close := "A/SSR_007_XV809_CFB",
                      reset := "Valves Data".R7_XV09.RESET OR "R7_DATA".R7.Reset,
                      intl := NOT "DI_INPUTS".R7_INPUTS_RUA.EMG_PB,
                      Mon_En := 1,
                      mon_sp := "Valves Data".R7_XV09.MON_TIME,
                      SEMI := "Valves Data".SEMI_AUTO.R7,
                      "open/close" => "A/SSR_007_XV809_CMD",
                      FAIL_TO_OPEN => "Valves Data".R7_VALVE_FAULT.XV09_FAIL_TO_OPEN,
                      FAIL_TO_CLOSE => "Valves Data".R7_VALVE_FAULT.XV09_FAIL_TO_CLOSE,
                      status => "Valves Data".R7_XV09.STATUS);
   END_IF;
END_REGION

REGION Network 76: R7_XV10
   RUNG wire#powerrail
      Contact( "AlwaysTRUE" )
      #valve_R7_XV10(reset := wire#w1, intl := wire#w2, "auto/manual" := "Valves Data"."A/M".R7, open_auto := "Valves Data".R7_XV10.CMD, open_man := "Valves Data".R7_XV10.MCMD, fbk_open := "A/SSR_007_XV401_OFB", fbk_close := "A/SSR_007_XV401_CFB", Mon_En := 1, mon_sp := "Valves Data".R7_XV10.MON_TIME, SEMI := "Valves Data".SEMI_AUTO.R7, SIM :=, "open/close" => "A/SSR_007_XV401_CMD", FAIL_TO_OPEN => "Valves Data".R7_VALVE_FAULT.XV010_FAIL_TO_OPEN, FAIL_TO_CLOSE => "Valves Data".R7_VALVE_FAULT.XV10_FAIL_TO_CLOSE, status => "Valves Data".R7_XV10.STATUS)
   END_RUNG
   RUNG wire#powerrail
      Contact( "Valves Data".R7_XV10.RESET )
   END_RUNG wire#w1
   RUNG wire#powerrail
      Contact( "R7_DATA".R7.Reset )
   END_RUNG wire#w1
   RUNG wire#powerrail
      I_Contact( "DI_INPUTS".R7_INPUTS_RUA.EMG_PB )
   END_RUNG wire#w2
   // the same network as SCL:
   IF "AlwaysTRUE" THEN
       #valve_R7_XV10("auto/manual" := "Valves Data"."A/M".R7,   // "valve"
                      open_auto := "Valves Data".R7_XV10.CMD,
                      open_man := "Valves Data".R7_XV10.MCMD,
                      fbk_open := "A/SSR_007_XV401_OFB",
                      fbk_close := "A/SSR_007_XV401_CFB",
                      reset := "Valves Data".R7_XV10.RESET OR "R7_DATA".R7.Reset,
                      intl := NOT "DI_INPUTS".R7_INPUTS_RUA.EMG_PB,
                      Mon_En := 1,
                      mon_sp := "Valves Data".R7_XV10.MON_TIME,
                      SEMI := "Valves Data".SEMI_AUTO.R7,
                      "open/close" => "A/SSR_007_XV401_CMD",
                      FAIL_TO_OPEN => "Valves Data".R7_VALVE_FAULT.XV010_FAIL_TO_OPEN,
                      FAIL_TO_CLOSE => "Valves Data".R7_VALVE_FAULT.XV10_FAIL_TO_CLOSE,
                      status => "Valves Data".R7_XV10.STATUS);
   END_IF;
END_REGION

REGION Network 77: ****REACTOR_08****
END_REGION

REGION Network 78: R8_XV01
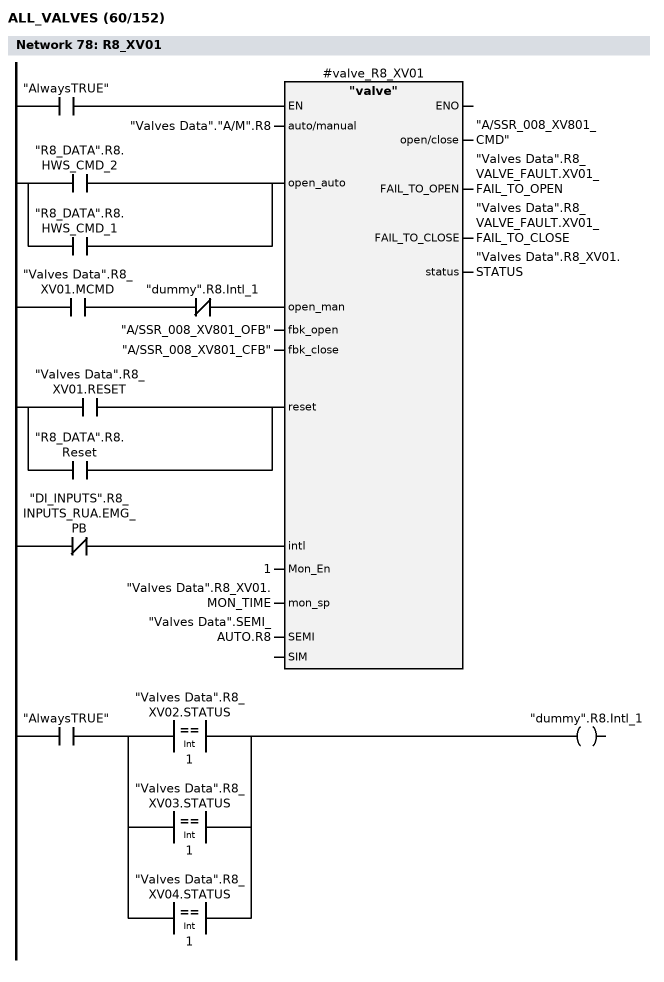
   RUNG wire#powerrail
      Contact( "AlwaysTRUE" )
      #valve_R8_XV01(open_auto := wire#w1, open_man := wire#w2, reset := wire#w3, intl := wire#w4, "auto/manual" := "Valves Data"."A/M".R8, fbk_open := "A/SSR_008_XV801_OFB", fbk_close := "A/SSR_008_XV801_CFB", Mon_En := 1, mon_sp := "Valves Data".R8_XV01.MON_TIME, SEMI := "Valves Data".SEMI_AUTO.R8, SIM :=, "open/close" => "A/SSR_008_XV801_CMD", FAIL_TO_OPEN => "Valves Data".R8_VALVE_FAULT.XV01_FAIL_TO_OPEN, FAIL_TO_CLOSE => "Valves Data".R8_VALVE_FAULT.XV01_FAIL_TO_CLOSE, status => "Valves Data".R8_XV01.STATUS)
   END_RUNG
   RUNG wire#powerrail
      Contact( "R8_DATA".R8.HWS_CMD_2 )
   END_RUNG wire#w1
   RUNG wire#powerrail
      Contact( "R8_DATA".R8.HWS_CMD_1 )
   END_RUNG wire#w1
   RUNG wire#powerrail
      Contact( "Valves Data".R8_XV01.MCMD )
      I_Contact( "dummy".R8.Intl_1 )
   END_RUNG wire#w2
   RUNG wire#powerrail
      Contact( "Valves Data".R8_XV01.RESET )
   END_RUNG wire#w3
   RUNG wire#powerrail
      Contact( "R8_DATA".R8.Reset )
   END_RUNG wire#w3
   RUNG wire#powerrail
      I_Contact( "DI_INPUTS".R8_INPUTS_RUA.EMG_PB )
   END_RUNG wire#w4
   RUNG wire#powerrail
      Contact( "AlwaysTRUE" )
      wire#w5
      { S7_Templates := "SrcType := Int" } EQ_Contact(in1 := "Valves Data".R8_XV02.STATUS, in2 := 1)
      wire#w6
      Coil( "dummy".R8.Intl_1 )
   END_RUNG
   RUNG wire#w5
      { S7_Templates := "SrcType := Int" } EQ_Contact(in1 := "Valves Data".R8_XV03.STATUS, in2 := 1)
   END_RUNG wire#w6
   RUNG wire#w5
      { S7_Templates := "SrcType := Int" } EQ_Contact(in1 := "Valves Data".R8_XV04.STATUS, in2 := 1)
   END_RUNG wire#w6
   // the same network as SCL:
   IF "AlwaysTRUE" THEN
       #valve_R8_XV01("auto/manual" := "Valves Data"."A/M".R8,   // "valve"
                      open_auto := "R8_DATA".R8.HWS_CMD_2 OR "R8_DATA".R8.HWS_CMD_1,
                      open_man := "Valves Data".R8_XV01.MCMD AND NOT "dummy".R8.Intl_1,
                      fbk_open := "A/SSR_008_XV801_OFB",
                      fbk_close := "A/SSR_008_XV801_CFB",
                      reset := "Valves Data".R8_XV01.RESET OR "R8_DATA".R8.Reset,
                      intl := NOT "DI_INPUTS".R8_INPUTS_RUA.EMG_PB,
                      Mon_En := 1,
                      mon_sp := "Valves Data".R8_XV01.MON_TIME,
                      SEMI := "Valves Data".SEMI_AUTO.R8,
                      "open/close" => "A/SSR_008_XV801_CMD",
                      FAIL_TO_OPEN => "Valves Data".R8_VALVE_FAULT.XV01_FAIL_TO_OPEN,
                      FAIL_TO_CLOSE => "Valves Data".R8_VALVE_FAULT.XV01_FAIL_TO_CLOSE,
                      status => "Valves Data".R8_XV01.STATUS);
   END_IF;
   "dummy".R8.Intl_1 := "AlwaysTRUE" AND (("Valves Data".R8_XV02.STATUS = 1) OR ("Valves Data".R8_XV03.STATUS = 1) OR ("Valves Data".R8_XV04.STATUS = 1));
END_REGION

REGION Network 79: R8_XV02
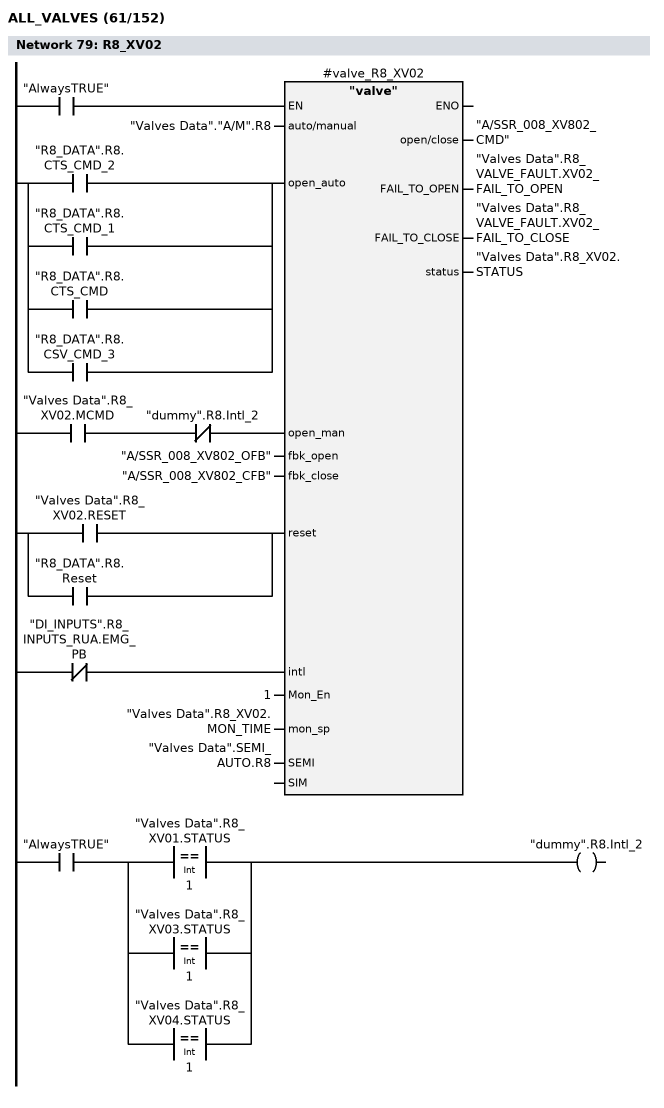
   RUNG wire#powerrail
      Contact( "AlwaysTRUE" )
      #valve_R8_XV02(open_auto := wire#w1, open_man := wire#w2, reset := wire#w3, intl := wire#w4, "auto/manual" := "Valves Data"."A/M".R8, fbk_open := "A/SSR_008_XV802_OFB", fbk_close := "A/SSR_008_XV802_CFB", Mon_En := 1, mon_sp := "Valves Data".R8_XV02.MON_TIME, SEMI := "Valves Data".SEMI_AUTO.R8, SIM :=, "open/close" => "A/SSR_008_XV802_CMD", FAIL_TO_OPEN => "Valves Data".R8_VALVE_FAULT.XV02_FAIL_TO_OPEN, FAIL_TO_CLOSE => "Valves Data".R8_VALVE_FAULT.XV02_FAIL_TO_CLOSE, status => "Valves Data".R8_XV02.STATUS)
   END_RUNG
   RUNG wire#powerrail
      Contact( "R8_DATA".R8.CTS_CMD_2 )
   END_RUNG wire#w1
   RUNG wire#powerrail
      Contact( "R8_DATA".R8.CTS_CMD_1 )
   END_RUNG wire#w1
   RUNG wire#powerrail
      Contact( "R8_DATA".R8.CTS_CMD )
   END_RUNG wire#w1
   RUNG wire#powerrail
      Contact( "R8_DATA".R8.CSV_CMD_3 )
   END_RUNG wire#w1
   RUNG wire#powerrail
      Contact( "Valves Data".R8_XV02.MCMD )
      I_Contact( "dummy".R8.Intl_2 )
   END_RUNG wire#w2
   RUNG wire#powerrail
      Contact( "Valves Data".R8_XV02.RESET )
   END_RUNG wire#w3
   RUNG wire#powerrail
      Contact( "R8_DATA".R8.Reset )
   END_RUNG wire#w3
   RUNG wire#powerrail
      I_Contact( "DI_INPUTS".R8_INPUTS_RUA.EMG_PB )
   END_RUNG wire#w4
   RUNG wire#powerrail
      Contact( "AlwaysTRUE" )
      wire#w5
      { S7_Templates := "SrcType := Int" } EQ_Contact(in1 := "Valves Data".R8_XV01.STATUS, in2 := 1)
      wire#w6
      Coil( "dummy".R8.Intl_2 )
   END_RUNG
   RUNG wire#w5
      { S7_Templates := "SrcType := Int" } EQ_Contact(in1 := "Valves Data".R8_XV03.STATUS, in2 := 1)
   END_RUNG wire#w6
   RUNG wire#w5
      { S7_Templates := "SrcType := Int" } EQ_Contact(in1 := "Valves Data".R8_XV04.STATUS, in2 := 1)
   END_RUNG wire#w6
   // the same network as SCL:
   IF "AlwaysTRUE" THEN
       #valve_R8_XV02("auto/manual" := "Valves Data"."A/M".R8,   // "valve"
                      open_auto := "R8_DATA".R8.CTS_CMD_2 OR "R8_DATA".R8.CTS_CMD_1 OR "R8_DATA".R8.CTS_CMD OR "R8_DATA".R8.CSV_CMD_3,
                      open_man := "Valves Data".R8_XV02.MCMD AND NOT "dummy".R8.Intl_2,
                      fbk_open := "A/SSR_008_XV802_OFB",
                      fbk_close := "A/SSR_008_XV802_CFB",
                      reset := "Valves Data".R8_XV02.RESET OR "R8_DATA".R8.Reset,
                      intl := NOT "DI_INPUTS".R8_INPUTS_RUA.EMG_PB,
                      Mon_En := 1,
                      mon_sp := "Valves Data".R8_XV02.MON_TIME,
                      SEMI := "Valves Data".SEMI_AUTO.R8,
                      "open/close" => "A/SSR_008_XV802_CMD",
                      FAIL_TO_OPEN => "Valves Data".R8_VALVE_FAULT.XV02_FAIL_TO_OPEN,
                      FAIL_TO_CLOSE => "Valves Data".R8_VALVE_FAULT.XV02_FAIL_TO_CLOSE,
                      status => "Valves Data".R8_XV02.STATUS);
   END_IF;
   "dummy".R8.Intl_2 := "AlwaysTRUE" AND (("Valves Data".R8_XV01.STATUS = 1) OR ("Valves Data".R8_XV03.STATUS = 1) OR ("Valves Data".R8_XV04.STATUS = 1));
END_REGION

REGION Network 80: R8_XV03
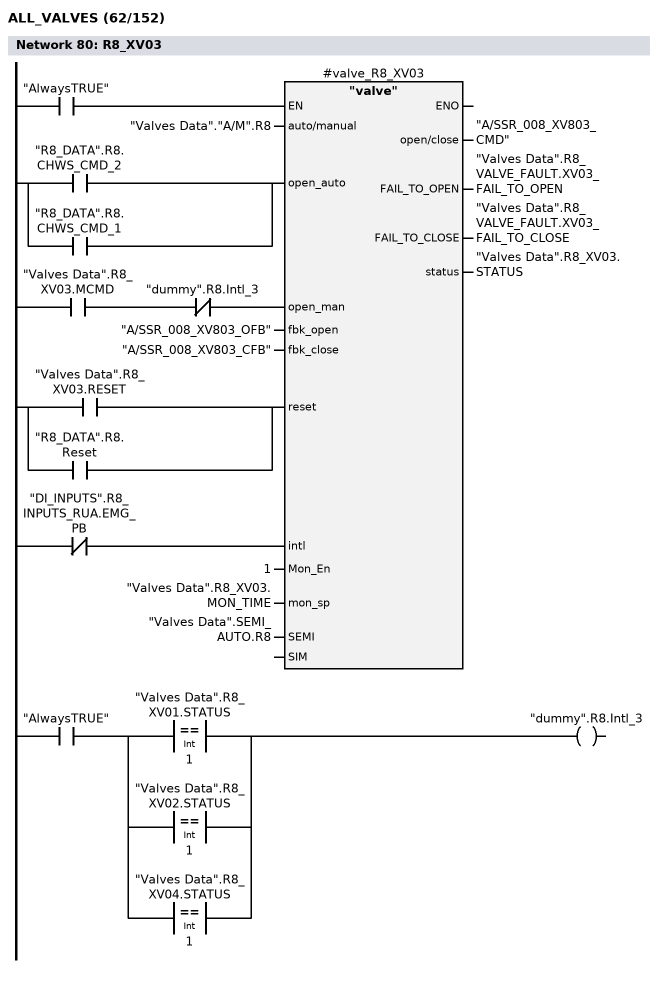
   RUNG wire#powerrail
      Contact( "AlwaysTRUE" )
      #valve_R8_XV03(open_auto := wire#w1, open_man := wire#w2, reset := wire#w3, intl := wire#w4, "auto/manual" := "Valves Data"."A/M".R8, fbk_open := "A/SSR_008_XV803_OFB", fbk_close := "A/SSR_008_XV803_CFB", Mon_En := 1, mon_sp := "Valves Data".R8_XV03.MON_TIME, SEMI := "Valves Data".SEMI_AUTO.R8, SIM :=, "open/close" => "A/SSR_008_XV803_CMD", FAIL_TO_OPEN => "Valves Data".R8_VALVE_FAULT.XV03_FAIL_TO_OPEN, FAIL_TO_CLOSE => "Valves Data".R8_VALVE_FAULT.XV03_FAIL_TO_CLOSE, status => "Valves Data".R8_XV03.STATUS)
   END_RUNG
   RUNG wire#powerrail
      Contact( "R8_DATA".R8.CHWS_CMD_2 )
   END_RUNG wire#w1
   RUNG wire#powerrail
      Contact( "R8_DATA".R8.CHWS_CMD_1 )
   END_RUNG wire#w1
   RUNG wire#powerrail
      Contact( "Valves Data".R8_XV03.MCMD )
      I_Contact( "dummy".R8.Intl_3 )
   END_RUNG wire#w2
   RUNG wire#powerrail
      Contact( "Valves Data".R8_XV03.RESET )
   END_RUNG wire#w3
   RUNG wire#powerrail
      Contact( "R8_DATA".R8.Reset )
   END_RUNG wire#w3
   RUNG wire#powerrail
      I_Contact( "DI_INPUTS".R8_INPUTS_RUA.EMG_PB )
   END_RUNG wire#w4
   RUNG wire#powerrail
      Contact( "AlwaysTRUE" )
      wire#w5
      { S7_Templates := "SrcType := Int" } EQ_Contact(in1 := "Valves Data".R8_XV01.STATUS, in2 := 1)
      wire#w6
      Coil( "dummy".R8.Intl_3 )
   END_RUNG
   RUNG wire#w5
      { S7_Templates := "SrcType := Int" } EQ_Contact(in1 := "Valves Data".R8_XV02.STATUS, in2 := 1)
   END_RUNG wire#w6
   RUNG wire#w5
      { S7_Templates := "SrcType := Int" } EQ_Contact(in1 := "Valves Data".R8_XV04.STATUS, in2 := 1)
   END_RUNG wire#w6
   // the same network as SCL:
   IF "AlwaysTRUE" THEN
       #valve_R8_XV03("auto/manual" := "Valves Data"."A/M".R8,   // "valve"
                      open_auto := "R8_DATA".R8.CHWS_CMD_2 OR "R8_DATA".R8.CHWS_CMD_1,
                      open_man := "Valves Data".R8_XV03.MCMD AND NOT "dummy".R8.Intl_3,
                      fbk_open := "A/SSR_008_XV803_OFB",
                      fbk_close := "A/SSR_008_XV803_CFB",
                      reset := "Valves Data".R8_XV03.RESET OR "R8_DATA".R8.Reset,
                      intl := NOT "DI_INPUTS".R8_INPUTS_RUA.EMG_PB,
                      Mon_En := 1,
                      mon_sp := "Valves Data".R8_XV03.MON_TIME,
                      SEMI := "Valves Data".SEMI_AUTO.R8,
                      "open/close" => "A/SSR_008_XV803_CMD",
                      FAIL_TO_OPEN => "Valves Data".R8_VALVE_FAULT.XV03_FAIL_TO_OPEN,
                      FAIL_TO_CLOSE => "Valves Data".R8_VALVE_FAULT.XV03_FAIL_TO_CLOSE,
                      status => "Valves Data".R8_XV03.STATUS);
   END_IF;
   "dummy".R8.Intl_3 := "AlwaysTRUE" AND (("Valves Data".R8_XV01.STATUS = 1) OR ("Valves Data".R8_XV02.STATUS = 1) OR ("Valves Data".R8_XV04.STATUS = 1));
END_REGION

REGION Network 81: R8_XV04
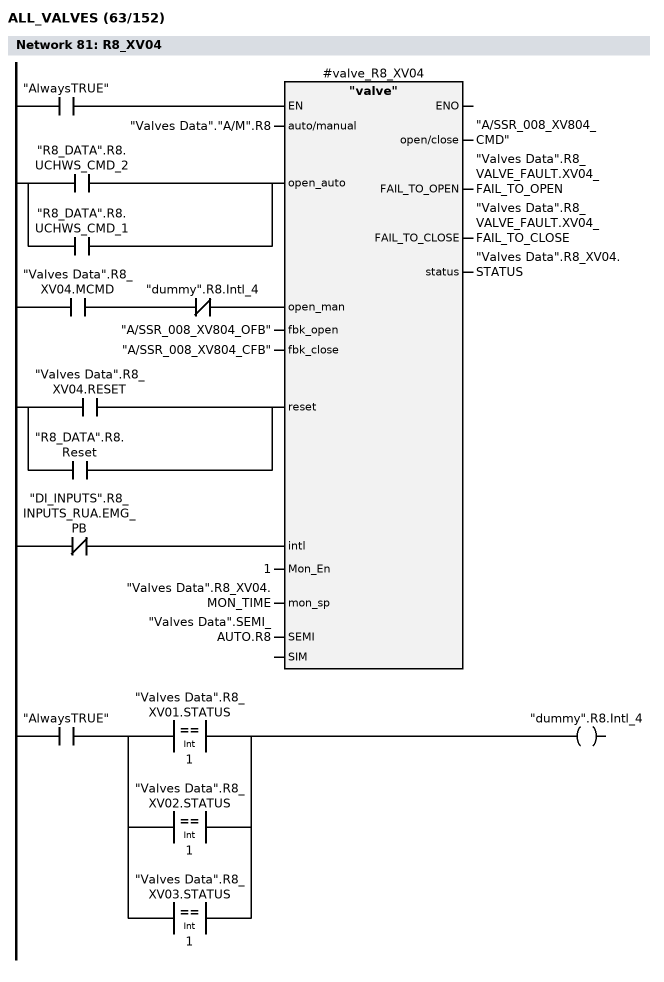
   RUNG wire#powerrail
      Contact( "AlwaysTRUE" )
      #valve_R8_XV04(open_auto := wire#w1, open_man := wire#w2, reset := wire#w3, intl := wire#w4, "auto/manual" := "Valves Data"."A/M".R8, fbk_open := "A/SSR_008_XV804_OFB", fbk_close := "A/SSR_008_XV804_CFB", Mon_En := 1, mon_sp := "Valves Data".R8_XV04.MON_TIME, SEMI := "Valves Data".SEMI_AUTO.R8, SIM :=, "open/close" => "A/SSR_008_XV804_CMD", FAIL_TO_OPEN => "Valves Data".R8_VALVE_FAULT.XV04_FAIL_TO_OPEN, FAIL_TO_CLOSE => "Valves Data".R8_VALVE_FAULT.XV04_FAIL_TO_CLOSE, status => "Valves Data".R8_XV04.STATUS)
   END_RUNG
   RUNG wire#powerrail
      Contact( "R8_DATA".R8.UCHWS_CMD_2 )
   END_RUNG wire#w1
   RUNG wire#powerrail
      Contact( "R8_DATA".R8.UCHWS_CMD_1 )
   END_RUNG wire#w1
   RUNG wire#powerrail
      Contact( "Valves Data".R8_XV04.MCMD )
      I_Contact( "dummy".R8.Intl_4 )
   END_RUNG wire#w2
   RUNG wire#powerrail
      Contact( "Valves Data".R8_XV04.RESET )
   END_RUNG wire#w3
   RUNG wire#powerrail
      Contact( "R8_DATA".R8.Reset )
   END_RUNG wire#w3
   RUNG wire#powerrail
      I_Contact( "DI_INPUTS".R8_INPUTS_RUA.EMG_PB )
   END_RUNG wire#w4
   RUNG wire#powerrail
      Contact( "AlwaysTRUE" )
      wire#w5
      { S7_Templates := "SrcType := Int" } EQ_Contact(in1 := "Valves Data".R8_XV01.STATUS, in2 := 1)
      wire#w6
      Coil( "dummy".R8.Intl_4 )
   END_RUNG
   RUNG wire#w5
      { S7_Templates := "SrcType := Int" } EQ_Contact(in1 := "Valves Data".R8_XV02.STATUS, in2 := 1)
   END_RUNG wire#w6
   RUNG wire#w5
      { S7_Templates := "SrcType := Int" } EQ_Contact(in1 := "Valves Data".R8_XV03.STATUS, in2 := 1)
   END_RUNG wire#w6
   // the same network as SCL:
   IF "AlwaysTRUE" THEN
       #valve_R8_XV04("auto/manual" := "Valves Data"."A/M".R8,   // "valve"
                      open_auto := "R8_DATA".R8.UCHWS_CMD_2 OR "R8_DATA".R8.UCHWS_CMD_1,
                      open_man := "Valves Data".R8_XV04.MCMD AND NOT "dummy".R8.Intl_4,
                      fbk_open := "A/SSR_008_XV804_OFB",
                      fbk_close := "A/SSR_008_XV804_CFB",
                      reset := "Valves Data".R8_XV04.RESET OR "R8_DATA".R8.Reset,
                      intl := NOT "DI_INPUTS".R8_INPUTS_RUA.EMG_PB,
                      Mon_En := 1,
                      mon_sp := "Valves Data".R8_XV04.MON_TIME,
                      SEMI := "Valves Data".SEMI_AUTO.R8,
                      "open/close" => "A/SSR_008_XV804_CMD",
                      FAIL_TO_OPEN => "Valves Data".R8_VALVE_FAULT.XV04_FAIL_TO_OPEN,
                      FAIL_TO_CLOSE => "Valves Data".R8_VALVE_FAULT.XV04_FAIL_TO_CLOSE,
                      status => "Valves Data".R8_XV04.STATUS);
   END_IF;
   "dummy".R8.Intl_4 := "AlwaysTRUE" AND (("Valves Data".R8_XV01.STATUS = 1) OR ("Valves Data".R8_XV02.STATUS = 1) OR ("Valves Data".R8_XV03.STATUS = 1));
END_REGION

REGION Network 82: R8_XV05
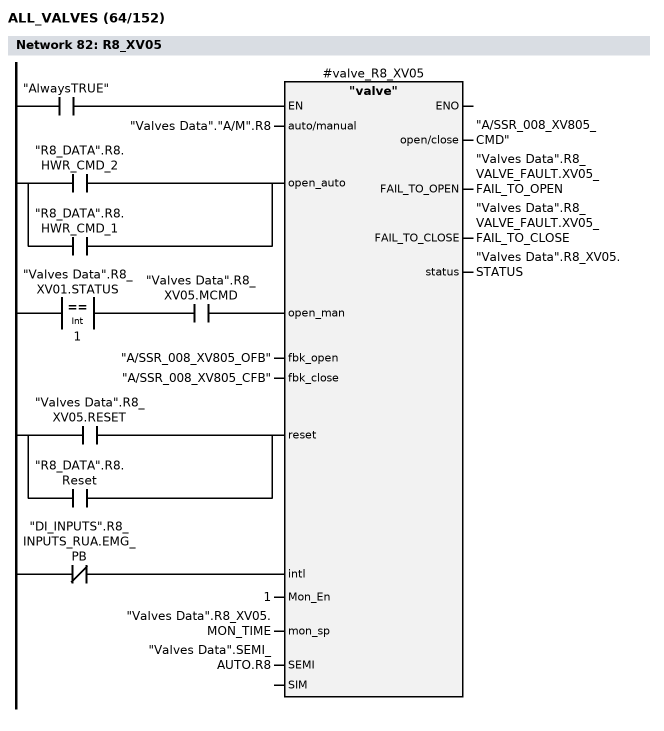
   RUNG wire#powerrail
      Contact( "AlwaysTRUE" )
      #valve_R8_XV05(open_auto := wire#w1, open_man := wire#w2, reset := wire#w3, intl := wire#w4, "auto/manual" := "Valves Data"."A/M".R8, fbk_open := "A/SSR_008_XV805_OFB", fbk_close := "A/SSR_008_XV805_CFB", Mon_En := 1, mon_sp := "Valves Data".R8_XV05.MON_TIME, SEMI := "Valves Data".SEMI_AUTO.R8, SIM :=, "open/close" => "A/SSR_008_XV805_CMD", FAIL_TO_OPEN => "Valves Data".R8_VALVE_FAULT.XV05_FAIL_TO_OPEN, FAIL_TO_CLOSE => "Valves Data".R8_VALVE_FAULT.XV05_FAIL_TO_CLOSE, status => "Valves Data".R8_XV05.STATUS)
   END_RUNG
   RUNG wire#powerrail
      Contact( "R8_DATA".R8.HWR_CMD_2 )
   END_RUNG wire#w1
   RUNG wire#powerrail
      Contact( "R8_DATA".R8.HWR_CMD_1 )
   END_RUNG wire#w1
   RUNG wire#powerrail
      { S7_Templates := "SrcType := Int" } EQ_Contact(in1 := "Valves Data".R8_XV01.STATUS, in2 := 1)
      Contact( "Valves Data".R8_XV05.MCMD )
   END_RUNG wire#w2
   RUNG wire#powerrail
      Contact( "Valves Data".R8_XV05.RESET )
   END_RUNG wire#w3
   RUNG wire#powerrail
      Contact( "R8_DATA".R8.Reset )
   END_RUNG wire#w3
   RUNG wire#powerrail
      I_Contact( "DI_INPUTS".R8_INPUTS_RUA.EMG_PB )
   END_RUNG wire#w4
   // the same network as SCL:
   IF "AlwaysTRUE" THEN
       #valve_R8_XV05("auto/manual" := "Valves Data"."A/M".R8,   // "valve"
                      open_auto := "R8_DATA".R8.HWR_CMD_2 OR "R8_DATA".R8.HWR_CMD_1,
                      open_man := ("Valves Data".R8_XV01.STATUS = 1) AND "Valves Data".R8_XV05.MCMD,
                      fbk_open := "A/SSR_008_XV805_OFB",
                      fbk_close := "A/SSR_008_XV805_CFB",
                      reset := "Valves Data".R8_XV05.RESET OR "R8_DATA".R8.Reset,
                      intl := NOT "DI_INPUTS".R8_INPUTS_RUA.EMG_PB,
                      Mon_En := 1,
                      mon_sp := "Valves Data".R8_XV05.MON_TIME,
                      SEMI := "Valves Data".SEMI_AUTO.R8,
                      "open/close" => "A/SSR_008_XV805_CMD",
                      FAIL_TO_OPEN => "Valves Data".R8_VALVE_FAULT.XV05_FAIL_TO_OPEN,
                      FAIL_TO_CLOSE => "Valves Data".R8_VALVE_FAULT.XV05_FAIL_TO_CLOSE,
                      status => "Valves Data".R8_XV05.STATUS);
   END_IF;
END_REGION

REGION Network 83: R8_XV06
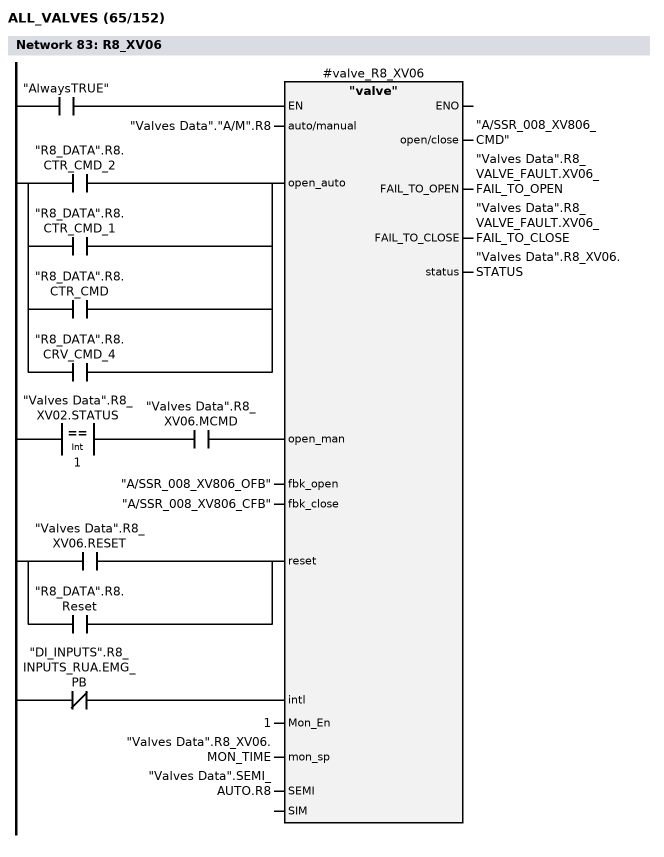
   RUNG wire#powerrail
      Contact( "AlwaysTRUE" )
      #valve_R8_XV06(open_auto := wire#w1, open_man := wire#w2, reset := wire#w3, intl := wire#w4, "auto/manual" := "Valves Data"."A/M".R8, fbk_open := "A/SSR_008_XV806_OFB", fbk_close := "A/SSR_008_XV806_CFB", Mon_En := 1, mon_sp := "Valves Data".R8_XV06.MON_TIME, SEMI := "Valves Data".SEMI_AUTO.R8, SIM :=, "open/close" => "A/SSR_008_XV806_CMD", FAIL_TO_OPEN => "Valves Data".R8_VALVE_FAULT.XV06_FAIL_TO_OPEN, FAIL_TO_CLOSE => "Valves Data".R8_VALVE_FAULT.XV06_FAIL_TO_CLOSE, status => "Valves Data".R8_XV06.STATUS)
   END_RUNG
   RUNG wire#powerrail
      Contact( "R8_DATA".R8.CTR_CMD_2 )
   END_RUNG wire#w1
   RUNG wire#powerrail
      Contact( "R8_DATA".R8.CTR_CMD_1 )
   END_RUNG wire#w1
   RUNG wire#powerrail
      Contact( "R8_DATA".R8.CTR_CMD )
   END_RUNG wire#w1
   RUNG wire#powerrail
      Contact( "R8_DATA".R8.CRV_CMD_4 )
   END_RUNG wire#w1
   RUNG wire#powerrail
      { S7_Templates := "SrcType := Int" } EQ_Contact(in1 := "Valves Data".R8_XV02.STATUS, in2 := 1)
      Contact( "Valves Data".R8_XV06.MCMD )
   END_RUNG wire#w2
   RUNG wire#powerrail
      Contact( "Valves Data".R8_XV06.RESET )
   END_RUNG wire#w3
   RUNG wire#powerrail
      Contact( "R8_DATA".R8.Reset )
   END_RUNG wire#w3
   RUNG wire#powerrail
      I_Contact( "DI_INPUTS".R8_INPUTS_RUA.EMG_PB )
   END_RUNG wire#w4
   // the same network as SCL:
   IF "AlwaysTRUE" THEN
       #valve_R8_XV06("auto/manual" := "Valves Data"."A/M".R8,   // "valve"
                      open_auto := "R8_DATA".R8.CTR_CMD_2 OR "R8_DATA".R8.CTR_CMD_1 OR "R8_DATA".R8.CTR_CMD OR "R8_DATA".R8.CRV_CMD_4,
                      open_man := ("Valves Data".R8_XV02.STATUS = 1) AND "Valves Data".R8_XV06.MCMD,
                      fbk_open := "A/SSR_008_XV806_OFB",
                      fbk_close := "A/SSR_008_XV806_CFB",
                      reset := "Valves Data".R8_XV06.RESET OR "R8_DATA".R8.Reset,
                      intl := NOT "DI_INPUTS".R8_INPUTS_RUA.EMG_PB,
                      Mon_En := 1,
                      mon_sp := "Valves Data".R8_XV06.MON_TIME,
                      SEMI := "Valves Data".SEMI_AUTO.R8,
                      "open/close" => "A/SSR_008_XV806_CMD",
                      FAIL_TO_OPEN => "Valves Data".R8_VALVE_FAULT.XV06_FAIL_TO_OPEN,
                      FAIL_TO_CLOSE => "Valves Data".R8_VALVE_FAULT.XV06_FAIL_TO_CLOSE,
                      status => "Valves Data".R8_XV06.STATUS);
   END_IF;
END_REGION

REGION Network 84: R8_XV07
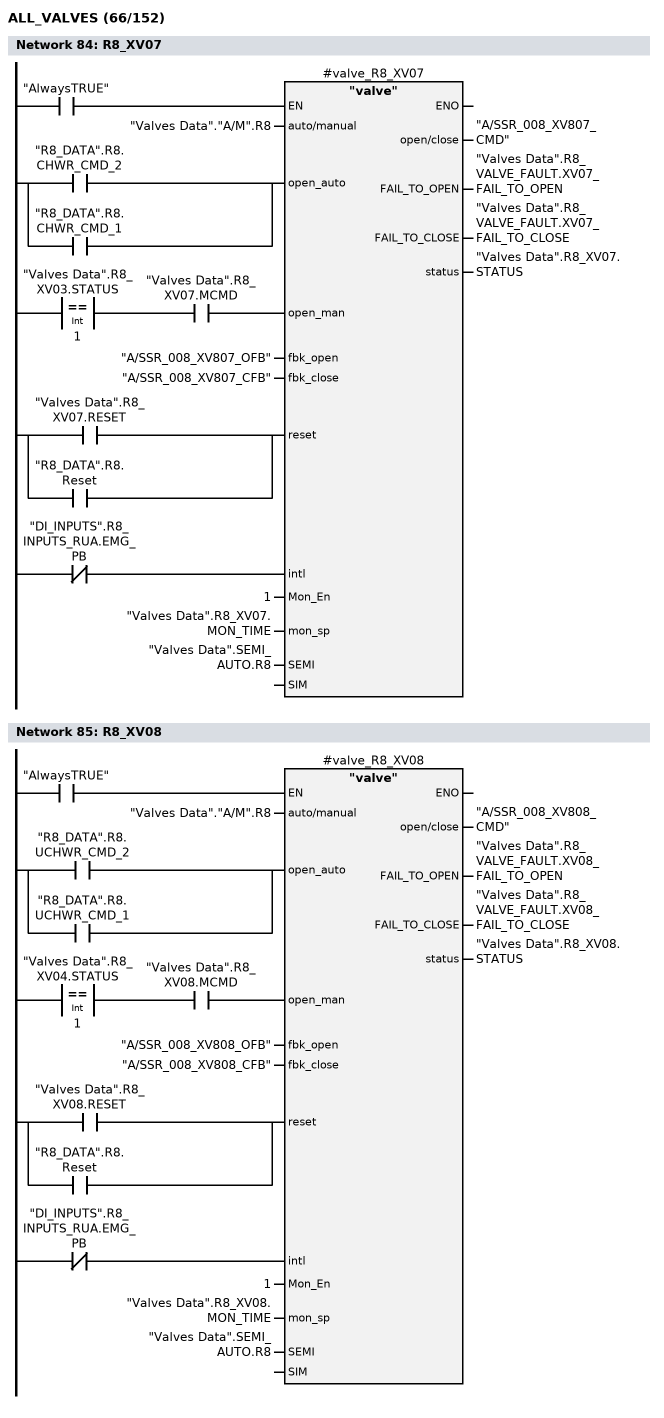
   RUNG wire#powerrail
      Contact( "AlwaysTRUE" )
      #valve_R8_XV07(open_auto := wire#w1, open_man := wire#w2, reset := wire#w3, intl := wire#w4, "auto/manual" := "Valves Data"."A/M".R8, fbk_open := "A/SSR_008_XV807_OFB", fbk_close := "A/SSR_008_XV807_CFB", Mon_En := 1, mon_sp := "Valves Data".R8_XV07.MON_TIME, SEMI := "Valves Data".SEMI_AUTO.R8, SIM :=, "open/close" => "A/SSR_008_XV807_CMD", FAIL_TO_OPEN => "Valves Data".R8_VALVE_FAULT.XV07_FAIL_TO_OPEN, FAIL_TO_CLOSE => "Valves Data".R8_VALVE_FAULT.XV07_FAIL_TO_CLOSE, status => "Valves Data".R8_XV07.STATUS)
   END_RUNG
   RUNG wire#powerrail
      Contact( "R8_DATA".R8.CHWR_CMD_2 )
   END_RUNG wire#w1
   RUNG wire#powerrail
      Contact( "R8_DATA".R8.CHWR_CMD_1 )
   END_RUNG wire#w1
   RUNG wire#powerrail
      { S7_Templates := "SrcType := Int" } EQ_Contact(in1 := "Valves Data".R8_XV03.STATUS, in2 := 1)
      Contact( "Valves Data".R8_XV07.MCMD )
   END_RUNG wire#w2
   RUNG wire#powerrail
      Contact( "Valves Data".R8_XV07.RESET )
   END_RUNG wire#w3
   RUNG wire#powerrail
      Contact( "R8_DATA".R8.Reset )
   END_RUNG wire#w3
   RUNG wire#powerrail
      I_Contact( "DI_INPUTS".R8_INPUTS_RUA.EMG_PB )
   END_RUNG wire#w4
   // the same network as SCL:
   IF "AlwaysTRUE" THEN
       #valve_R8_XV07("auto/manual" := "Valves Data"."A/M".R8,   // "valve"
                      open_auto := "R8_DATA".R8.CHWR_CMD_2 OR "R8_DATA".R8.CHWR_CMD_1,
                      open_man := ("Valves Data".R8_XV03.STATUS = 1) AND "Valves Data".R8_XV07.MCMD,
                      fbk_open := "A/SSR_008_XV807_OFB",
                      fbk_close := "A/SSR_008_XV807_CFB",
                      reset := "Valves Data".R8_XV07.RESET OR "R8_DATA".R8.Reset,
                      intl := NOT "DI_INPUTS".R8_INPUTS_RUA.EMG_PB,
                      Mon_En := 1,
                      mon_sp := "Valves Data".R8_XV07.MON_TIME,
                      SEMI := "Valves Data".SEMI_AUTO.R8,
                      "open/close" => "A/SSR_008_XV807_CMD",
                      FAIL_TO_OPEN => "Valves Data".R8_VALVE_FAULT.XV07_FAIL_TO_OPEN,
                      FAIL_TO_CLOSE => "Valves Data".R8_VALVE_FAULT.XV07_FAIL_TO_CLOSE,
                      status => "Valves Data".R8_XV07.STATUS);
   END_IF;
END_REGION

REGION Network 85: R8_XV08
   RUNG wire#powerrail
      Contact( "AlwaysTRUE" )
      #valve_R8_XV08(open_auto := wire#w1, open_man := wire#w2, reset := wire#w3, intl := wire#w4, "auto/manual" := "Valves Data"."A/M".R8, fbk_open := "A/SSR_008_XV808_OFB", fbk_close := "A/SSR_008_XV808_CFB", Mon_En := 1, mon_sp := "Valves Data".R8_XV08.MON_TIME, SEMI := "Valves Data".SEMI_AUTO.R8, SIM :=, "open/close" => "A/SSR_008_XV808_CMD", FAIL_TO_OPEN => "Valves Data".R8_VALVE_FAULT.XV08_FAIL_TO_OPEN, FAIL_TO_CLOSE => "Valves Data".R8_VALVE_FAULT.XV08_FAIL_TO_CLOSE, status => "Valves Data".R8_XV08.STATUS)
   END_RUNG
   RUNG wire#powerrail
      Contact( "R8_DATA".R8.UCHWR_CMD_2 )
   END_RUNG wire#w1
   RUNG wire#powerrail
      Contact( "R8_DATA".R8.UCHWR_CMD_1 )
   END_RUNG wire#w1
   RUNG wire#powerrail
      { S7_Templates := "SrcType := Int" } EQ_Contact(in1 := "Valves Data".R8_XV04.STATUS, in2 := 1)
      Contact( "Valves Data".R8_XV08.MCMD )
   END_RUNG wire#w2
   RUNG wire#powerrail
      Contact( "Valves Data".R8_XV08.RESET )
   END_RUNG wire#w3
   RUNG wire#powerrail
      Contact( "R8_DATA".R8.Reset )
   END_RUNG wire#w3
   RUNG wire#powerrail
      I_Contact( "DI_INPUTS".R8_INPUTS_RUA.EMG_PB )
   END_RUNG wire#w4
   // the same network as SCL:
   IF "AlwaysTRUE" THEN
       #valve_R8_XV08("auto/manual" := "Valves Data"."A/M".R8,   // "valve"
                      open_auto := "R8_DATA".R8.UCHWR_CMD_2 OR "R8_DATA".R8.UCHWR_CMD_1,
                      open_man := ("Valves Data".R8_XV04.STATUS = 1) AND "Valves Data".R8_XV08.MCMD,
                      fbk_open := "A/SSR_008_XV808_OFB",
                      fbk_close := "A/SSR_008_XV808_CFB",
                      reset := "Valves Data".R8_XV08.RESET OR "R8_DATA".R8.Reset,
                      intl := NOT "DI_INPUTS".R8_INPUTS_RUA.EMG_PB,
                      Mon_En := 1,
                      mon_sp := "Valves Data".R8_XV08.MON_TIME,
                      SEMI := "Valves Data".SEMI_AUTO.R8,
                      "open/close" => "A/SSR_008_XV808_CMD",
                      FAIL_TO_OPEN => "Valves Data".R8_VALVE_FAULT.XV08_FAIL_TO_OPEN,
                      FAIL_TO_CLOSE => "Valves Data".R8_VALVE_FAULT.XV08_FAIL_TO_CLOSE,
                      status => "Valves Data".R8_XV08.STATUS);
   END_IF;
END_REGION

REGION Network 86: R8_XV09
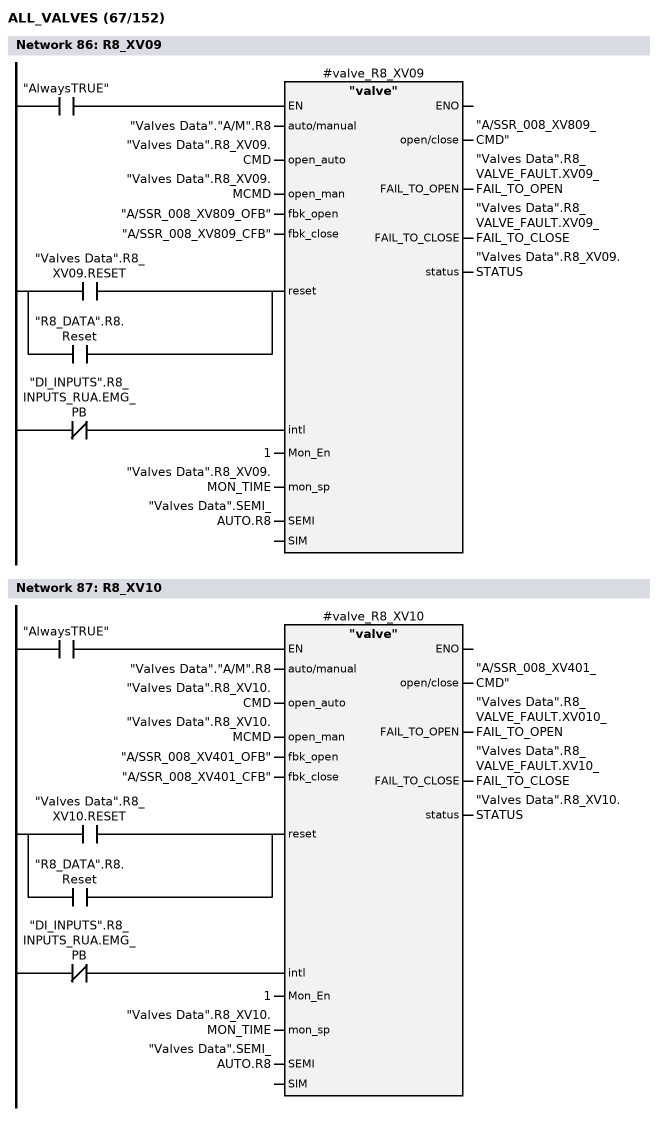
   RUNG wire#powerrail
      Contact( "AlwaysTRUE" )
      #valve_R8_XV09(reset := wire#w1, intl := wire#w2, "auto/manual" := "Valves Data"."A/M".R8, open_auto := "Valves Data".R8_XV09.CMD, open_man := "Valves Data".R8_XV09.MCMD, fbk_open := "A/SSR_008_XV809_OFB", fbk_close := "A/SSR_008_XV809_CFB", Mon_En := 1, mon_sp := "Valves Data".R8_XV09.MON_TIME, SEMI := "Valves Data".SEMI_AUTO.R8, SIM :=, "open/close" => "A/SSR_008_XV809_CMD", FAIL_TO_OPEN => "Valves Data".R8_VALVE_FAULT.XV09_FAIL_TO_OPEN, FAIL_TO_CLOSE => "Valves Data".R8_VALVE_FAULT.XV09_FAIL_TO_CLOSE, status => "Valves Data".R8_XV09.STATUS)
   END_RUNG
   RUNG wire#powerrail
      Contact( "Valves Data".R8_XV09.RESET )
   END_RUNG wire#w1
   RUNG wire#powerrail
      Contact( "R8_DATA".R8.Reset )
   END_RUNG wire#w1
   RUNG wire#powerrail
      I_Contact( "DI_INPUTS".R8_INPUTS_RUA.EMG_PB )
   END_RUNG wire#w2
   // the same network as SCL:
   IF "AlwaysTRUE" THEN
       #valve_R8_XV09("auto/manual" := "Valves Data"."A/M".R8,   // "valve"
                      open_auto := "Valves Data".R8_XV09.CMD,
                      open_man := "Valves Data".R8_XV09.MCMD,
                      fbk_open := "A/SSR_008_XV809_OFB",
                      fbk_close := "A/SSR_008_XV809_CFB",
                      reset := "Valves Data".R8_XV09.RESET OR "R8_DATA".R8.Reset,
                      intl := NOT "DI_INPUTS".R8_INPUTS_RUA.EMG_PB,
                      Mon_En := 1,
                      mon_sp := "Valves Data".R8_XV09.MON_TIME,
                      SEMI := "Valves Data".SEMI_AUTO.R8,
                      "open/close" => "A/SSR_008_XV809_CMD",
                      FAIL_TO_OPEN => "Valves Data".R8_VALVE_FAULT.XV09_FAIL_TO_OPEN,
                      FAIL_TO_CLOSE => "Valves Data".R8_VALVE_FAULT.XV09_FAIL_TO_CLOSE,
                      status => "Valves Data".R8_XV09.STATUS);
   END_IF;
END_REGION

REGION Network 87: R8_XV10
   RUNG wire#powerrail
      Contact( "AlwaysTRUE" )
      #valve_R8_XV10(reset := wire#w1, intl := wire#w2, "auto/manual" := "Valves Data"."A/M".R8, open_auto := "Valves Data".R8_XV10.CMD, open_man := "Valves Data".R8_XV10.MCMD, fbk_open := "A/SSR_008_XV401_OFB", fbk_close := "A/SSR_008_XV401_CFB", Mon_En := 1, mon_sp := "Valves Data".R8_XV10.MON_TIME, SEMI := "Valves Data".SEMI_AUTO.R8, SIM :=, "open/close" => "A/SSR_008_XV401_CMD", FAIL_TO_OPEN => "Valves Data".R8_VALVE_FAULT.XV010_FAIL_TO_OPEN, FAIL_TO_CLOSE => "Valves Data".R8_VALVE_FAULT.XV10_FAIL_TO_CLOSE, status => "Valves Data".R8_XV10.STATUS)
   END_RUNG
   RUNG wire#powerrail
      Contact( "Valves Data".R8_XV10.RESET )
   END_RUNG wire#w1
   RUNG wire#powerrail
      Contact( "R8_DATA".R8.Reset )
   END_RUNG wire#w1
   RUNG wire#powerrail
      I_Contact( "DI_INPUTS".R8_INPUTS_RUA.EMG_PB )
   END_RUNG wire#w2
   // the same network as SCL:
   IF "AlwaysTRUE" THEN
       #valve_R8_XV10("auto/manual" := "Valves Data"."A/M".R8,   // "valve"
                      open_auto := "Valves Data".R8_XV10.CMD,
                      open_man := "Valves Data".R8_XV10.MCMD,
                      fbk_open := "A/SSR_008_XV401_OFB",
                      fbk_close := "A/SSR_008_XV401_CFB",
                      reset := "Valves Data".R8_XV10.RESET OR "R8_DATA".R8.Reset,
                      intl := NOT "DI_INPUTS".R8_INPUTS_RUA.EMG_PB,
                      Mon_En := 1,
                      mon_sp := "Valves Data".R8_XV10.MON_TIME,
                      SEMI := "Valves Data".SEMI_AUTO.R8,
                      "open/close" => "A/SSR_008_XV401_CMD",
                      FAIL_TO_OPEN => "Valves Data".R8_VALVE_FAULT.XV010_FAIL_TO_OPEN,
                      FAIL_TO_CLOSE => "Valves Data".R8_VALVE_FAULT.XV10_FAIL_TO_CLOSE,
                      status => "Valves Data".R8_XV10.STATUS);
   END_IF;
END_REGION

REGION Network 88: ****REACTOR_09****
END_REGION

REGION Network 89: R9_XV01
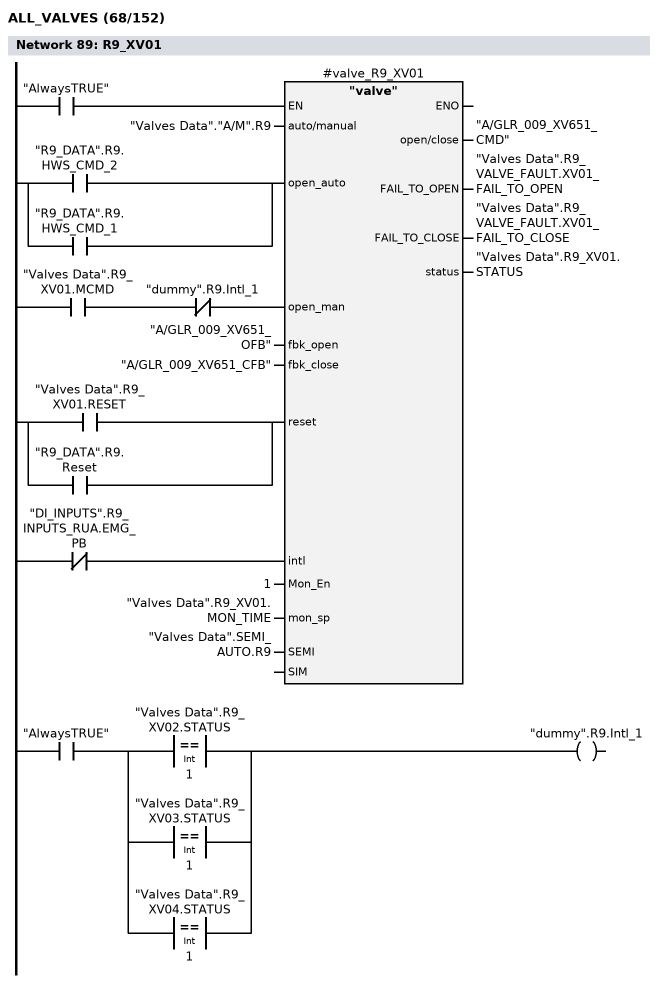
   RUNG wire#powerrail
      Contact( "AlwaysTRUE" )
      #valve_R9_XV01(open_auto := wire#w1, open_man := wire#w2, reset := wire#w3, intl := wire#w4, "auto/manual" := "Valves Data"."A/M".R9, fbk_open := "A/GLR_009_XV651_OFB", fbk_close := "A/GLR_009_XV651_CFB", Mon_En := 1, mon_sp := "Valves Data".R9_XV01.MON_TIME, SEMI := "Valves Data".SEMI_AUTO.R9, SIM :=, "open/close" => "A/GLR_009_XV651_CMD", FAIL_TO_OPEN => "Valves Data".R9_VALVE_FAULT.XV01_FAIL_TO_OPEN, FAIL_TO_CLOSE => "Valves Data".R9_VALVE_FAULT.XV01_FAIL_TO_CLOSE, status => "Valves Data".R9_XV01.STATUS)
   END_RUNG
   RUNG wire#powerrail
      Contact( "R9_DATA".R9.HWS_CMD_2 )
   END_RUNG wire#w1
   RUNG wire#powerrail
      Contact( "R9_DATA".R9.HWS_CMD_1 )
   END_RUNG wire#w1
   RUNG wire#powerrail
      Contact( "Valves Data".R9_XV01.MCMD )
      I_Contact( "dummy".R9.Intl_1 )
   END_RUNG wire#w2
   RUNG wire#powerrail
      Contact( "Valves Data".R9_XV01.RESET )
   END_RUNG wire#w3
   RUNG wire#powerrail
      Contact( "R9_DATA".R9.Reset )
   END_RUNG wire#w3
   RUNG wire#powerrail
      I_Contact( "DI_INPUTS".R9_INPUTS_RUA.EMG_PB )
   END_RUNG wire#w4
   RUNG wire#powerrail
      Contact( "AlwaysTRUE" )
      wire#w5
      { S7_Templates := "SrcType := Int" } EQ_Contact(in1 := "Valves Data".R9_XV02.STATUS, in2 := 1)
      wire#w6
      Coil( "dummy".R9.Intl_1 )
   END_RUNG
   RUNG wire#w5
      { S7_Templates := "SrcType := Int" } EQ_Contact(in1 := "Valves Data".R9_XV03.STATUS, in2 := 1)
   END_RUNG wire#w6
   RUNG wire#w5
      { S7_Templates := "SrcType := Int" } EQ_Contact(in1 := "Valves Data".R9_XV04.STATUS, in2 := 1)
   END_RUNG wire#w6
   // the same network as SCL:
   IF "AlwaysTRUE" THEN
       #valve_R9_XV01("auto/manual" := "Valves Data"."A/M".R9,   // "valve"
                      open_auto := "R9_DATA".R9.HWS_CMD_2 OR "R9_DATA".R9.HWS_CMD_1,
                      open_man := "Valves Data".R9_XV01.MCMD AND NOT "dummy".R9.Intl_1,
                      fbk_open := "A/GLR_009_XV651_OFB",
                      fbk_close := "A/GLR_009_XV651_CFB",
                      reset := "Valves Data".R9_XV01.RESET OR "R9_DATA".R9.Reset,
                      intl := NOT "DI_INPUTS".R9_INPUTS_RUA.EMG_PB,
                      Mon_En := 1,
                      mon_sp := "Valves Data".R9_XV01.MON_TIME,
                      SEMI := "Valves Data".SEMI_AUTO.R9,
                      "open/close" => "A/GLR_009_XV651_CMD",
                      FAIL_TO_OPEN => "Valves Data".R9_VALVE_FAULT.XV01_FAIL_TO_OPEN,
                      FAIL_TO_CLOSE => "Valves Data".R9_VALVE_FAULT.XV01_FAIL_TO_CLOSE,
                      status => "Valves Data".R9_XV01.STATUS);
   END_IF;
   "dummy".R9.Intl_1 := "AlwaysTRUE" AND (("Valves Data".R9_XV02.STATUS = 1) OR ("Valves Data".R9_XV03.STATUS = 1) OR ("Valves Data".R9_XV04.STATUS = 1));
END_REGION

REGION Network 90: R9_XV02
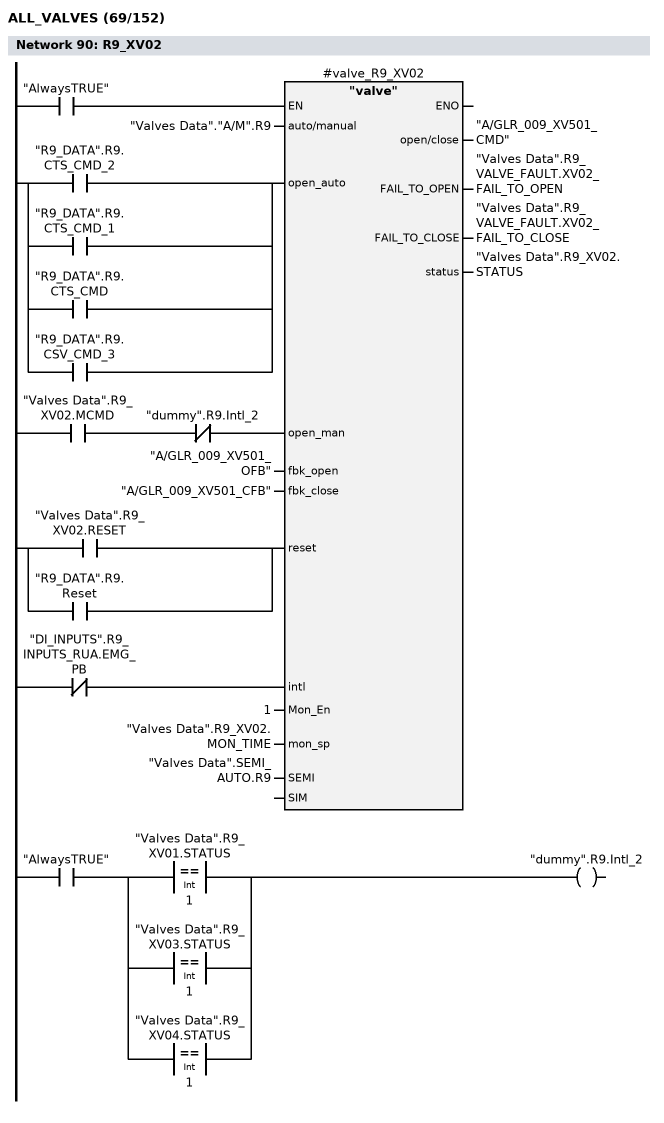
   RUNG wire#powerrail
      Contact( "AlwaysTRUE" )
      #valve_R9_XV02(open_auto := wire#w1, open_man := wire#w2, reset := wire#w3, intl := wire#w4, "auto/manual" := "Valves Data"."A/M".R9, fbk_open := "A/GLR_009_XV501_OFB", fbk_close := "A/GLR_009_XV501_CFB", Mon_En := 1, mon_sp := "Valves Data".R9_XV02.MON_TIME, SEMI := "Valves Data".SEMI_AUTO.R9, SIM :=, "open/close" => "A/GLR_009_XV501_CMD", FAIL_TO_OPEN => "Valves Data".R9_VALVE_FAULT.XV02_FAIL_TO_OPEN, FAIL_TO_CLOSE => "Valves Data".R9_VALVE_FAULT.XV02_FAIL_TO_CLOSE, status => "Valves Data".R9_XV02.STATUS)
   END_RUNG
   RUNG wire#powerrail
      Contact( "R9_DATA".R9.CTS_CMD_2 )
   END_RUNG wire#w1
   RUNG wire#powerrail
      Contact( "R9_DATA".R9.CTS_CMD_1 )
   END_RUNG wire#w1
   RUNG wire#powerrail
      Contact( "R9_DATA".R9.CTS_CMD )
   END_RUNG wire#w1
   RUNG wire#powerrail
      Contact( "R9_DATA".R9.CSV_CMD_3 )
   END_RUNG wire#w1
   RUNG wire#powerrail
      Contact( "Valves Data".R9_XV02.MCMD )
      I_Contact( "dummy".R9.Intl_2 )
   END_RUNG wire#w2
   RUNG wire#powerrail
      Contact( "Valves Data".R9_XV02.RESET )
   END_RUNG wire#w3
   RUNG wire#powerrail
      Contact( "R9_DATA".R9.Reset )
   END_RUNG wire#w3
   RUNG wire#powerrail
      I_Contact( "DI_INPUTS".R9_INPUTS_RUA.EMG_PB )
   END_RUNG wire#w4
   RUNG wire#powerrail
      Contact( "AlwaysTRUE" )
      wire#w5
      { S7_Templates := "SrcType := Int" } EQ_Contact(in1 := "Valves Data".R9_XV01.STATUS, in2 := 1)
      wire#w6
      Coil( "dummy".R9.Intl_2 )
   END_RUNG
   RUNG wire#w5
      { S7_Templates := "SrcType := Int" } EQ_Contact(in1 := "Valves Data".R9_XV03.STATUS, in2 := 1)
   END_RUNG wire#w6
   RUNG wire#w5
      { S7_Templates := "SrcType := Int" } EQ_Contact(in1 := "Valves Data".R9_XV04.STATUS, in2 := 1)
   END_RUNG wire#w6
   // the same network as SCL:
   IF "AlwaysTRUE" THEN
       #valve_R9_XV02("auto/manual" := "Valves Data"."A/M".R9,   // "valve"
                      open_auto := "R9_DATA".R9.CTS_CMD_2 OR "R9_DATA".R9.CTS_CMD_1 OR "R9_DATA".R9.CTS_CMD OR "R9_DATA".R9.CSV_CMD_3,
                      open_man := "Valves Data".R9_XV02.MCMD AND NOT "dummy".R9.Intl_2,
                      fbk_open := "A/GLR_009_XV501_OFB",
                      fbk_close := "A/GLR_009_XV501_CFB",
                      reset := "Valves Data".R9_XV02.RESET OR "R9_DATA".R9.Reset,
                      intl := NOT "DI_INPUTS".R9_INPUTS_RUA.EMG_PB,
                      Mon_En := 1,
                      mon_sp := "Valves Data".R9_XV02.MON_TIME,
                      SEMI := "Valves Data".SEMI_AUTO.R9,
                      "open/close" => "A/GLR_009_XV501_CMD",
                      FAIL_TO_OPEN => "Valves Data".R9_VALVE_FAULT.XV02_FAIL_TO_OPEN,
                      FAIL_TO_CLOSE => "Valves Data".R9_VALVE_FAULT.XV02_FAIL_TO_CLOSE,
                      status => "Valves Data".R9_XV02.STATUS);
   END_IF;
   "dummy".R9.Intl_2 := "AlwaysTRUE" AND (("Valves Data".R9_XV01.STATUS = 1) OR ("Valves Data".R9_XV03.STATUS = 1) OR ("Valves Data".R9_XV04.STATUS = 1));
END_REGION

REGION Network 91: R9_XV03
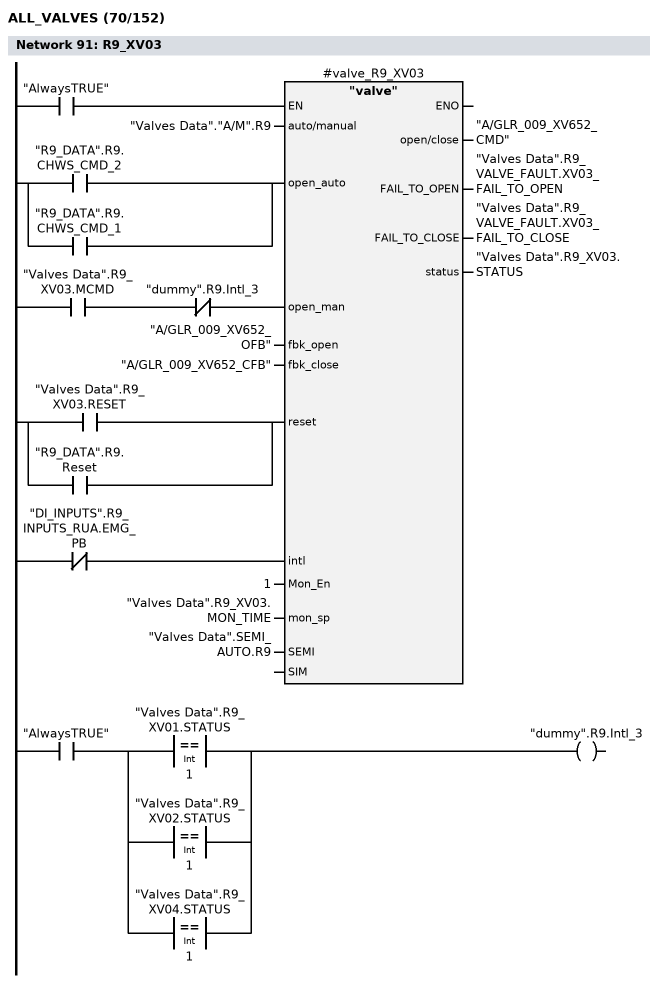
   RUNG wire#powerrail
      Contact( "AlwaysTRUE" )
      #valve_R9_XV03(open_auto := wire#w1, open_man := wire#w2, reset := wire#w3, intl := wire#w4, "auto/manual" := "Valves Data"."A/M".R9, fbk_open := "A/GLR_009_XV652_OFB", fbk_close := "A/GLR_009_XV652_CFB", Mon_En := 1, mon_sp := "Valves Data".R9_XV03.MON_TIME, SEMI := "Valves Data".SEMI_AUTO.R9, SIM :=, "open/close" => "A/GLR_009_XV652_CMD", FAIL_TO_OPEN => "Valves Data".R9_VALVE_FAULT.XV03_FAIL_TO_OPEN, FAIL_TO_CLOSE => "Valves Data".R9_VALVE_FAULT.XV03_FAIL_TO_CLOSE, status => "Valves Data".R9_XV03.STATUS)
   END_RUNG
   RUNG wire#powerrail
      Contact( "R9_DATA".R9.CHWS_CMD_2 )
   END_RUNG wire#w1
   RUNG wire#powerrail
      Contact( "R9_DATA".R9.CHWS_CMD_1 )
   END_RUNG wire#w1
   RUNG wire#powerrail
      Contact( "Valves Data".R9_XV03.MCMD )
      I_Contact( "dummy".R9.Intl_3 )
   END_RUNG wire#w2
   RUNG wire#powerrail
      Contact( "Valves Data".R9_XV03.RESET )
   END_RUNG wire#w3
   RUNG wire#powerrail
      Contact( "R9_DATA".R9.Reset )
   END_RUNG wire#w3
   RUNG wire#powerrail
      I_Contact( "DI_INPUTS".R9_INPUTS_RUA.EMG_PB )
   END_RUNG wire#w4
   RUNG wire#powerrail
      Contact( "AlwaysTRUE" )
      wire#w5
      { S7_Templates := "SrcType := Int" } EQ_Contact(in1 := "Valves Data".R9_XV01.STATUS, in2 := 1)
      wire#w6
      Coil( "dummy".R9.Intl_3 )
   END_RUNG
   RUNG wire#w5
      { S7_Templates := "SrcType := Int" } EQ_Contact(in1 := "Valves Data".R9_XV02.STATUS, in2 := 1)
   END_RUNG wire#w6
   RUNG wire#w5
      { S7_Templates := "SrcType := Int" } EQ_Contact(in1 := "Valves Data".R9_XV04.STATUS, in2 := 1)
   END_RUNG wire#w6
   // the same network as SCL:
   IF "AlwaysTRUE" THEN
       #valve_R9_XV03("auto/manual" := "Valves Data"."A/M".R9,   // "valve"
                      open_auto := "R9_DATA".R9.CHWS_CMD_2 OR "R9_DATA".R9.CHWS_CMD_1,
                      open_man := "Valves Data".R9_XV03.MCMD AND NOT "dummy".R9.Intl_3,
                      fbk_open := "A/GLR_009_XV652_OFB",
                      fbk_close := "A/GLR_009_XV652_CFB",
                      reset := "Valves Data".R9_XV03.RESET OR "R9_DATA".R9.Reset,
                      intl := NOT "DI_INPUTS".R9_INPUTS_RUA.EMG_PB,
                      Mon_En := 1,
                      mon_sp := "Valves Data".R9_XV03.MON_TIME,
                      SEMI := "Valves Data".SEMI_AUTO.R9,
                      "open/close" => "A/GLR_009_XV652_CMD",
                      FAIL_TO_OPEN => "Valves Data".R9_VALVE_FAULT.XV03_FAIL_TO_OPEN,
                      FAIL_TO_CLOSE => "Valves Data".R9_VALVE_FAULT.XV03_FAIL_TO_CLOSE,
                      status => "Valves Data".R9_XV03.STATUS);
   END_IF;
   "dummy".R9.Intl_3 := "AlwaysTRUE" AND (("Valves Data".R9_XV01.STATUS = 1) OR ("Valves Data".R9_XV02.STATUS = 1) OR ("Valves Data".R9_XV04.STATUS = 1));
END_REGION

REGION Network 92: R9_XV04
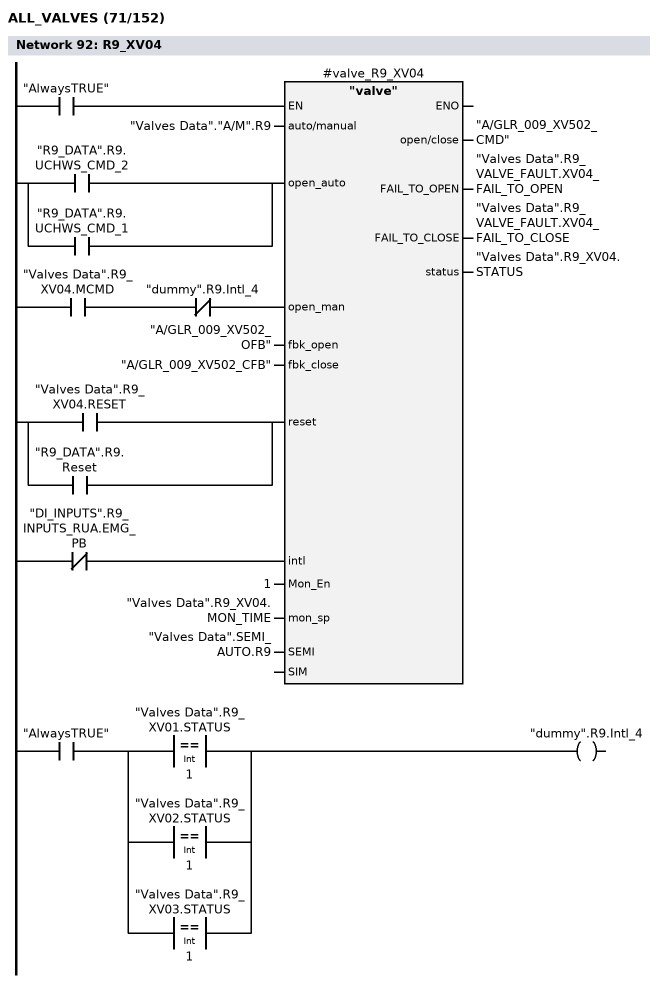
   RUNG wire#powerrail
      Contact( "AlwaysTRUE" )
      #valve_R9_XV04(open_auto := wire#w1, open_man := wire#w2, reset := wire#w3, intl := wire#w4, "auto/manual" := "Valves Data"."A/M".R9, fbk_open := "A/GLR_009_XV502_OFB", fbk_close := "A/GLR_009_XV502_CFB", Mon_En := 1, mon_sp := "Valves Data".R9_XV04.MON_TIME, SEMI := "Valves Data".SEMI_AUTO.R9, SIM :=, "open/close" => "A/GLR_009_XV502_CMD", FAIL_TO_OPEN => "Valves Data".R9_VALVE_FAULT.XV04_FAIL_TO_OPEN, FAIL_TO_CLOSE => "Valves Data".R9_VALVE_FAULT.XV04_FAIL_TO_CLOSE, status => "Valves Data".R9_XV04.STATUS)
   END_RUNG
   RUNG wire#powerrail
      Contact( "R9_DATA".R9.UCHWS_CMD_2 )
   END_RUNG wire#w1
   RUNG wire#powerrail
      Contact( "R9_DATA".R9.UCHWS_CMD_1 )
   END_RUNG wire#w1
   RUNG wire#powerrail
      Contact( "Valves Data".R9_XV04.MCMD )
      I_Contact( "dummy".R9.Intl_4 )
   END_RUNG wire#w2
   RUNG wire#powerrail
      Contact( "Valves Data".R9_XV04.RESET )
   END_RUNG wire#w3
   RUNG wire#powerrail
      Contact( "R9_DATA".R9.Reset )
   END_RUNG wire#w3
   RUNG wire#powerrail
      I_Contact( "DI_INPUTS".R9_INPUTS_RUA.EMG_PB )
   END_RUNG wire#w4
   RUNG wire#powerrail
      Contact( "AlwaysTRUE" )
      wire#w5
      { S7_Templates := "SrcType := Int" } EQ_Contact(in1 := "Valves Data".R9_XV01.STATUS, in2 := 1)
      wire#w6
      Coil( "dummy".R9.Intl_4 )
   END_RUNG
   RUNG wire#w5
      { S7_Templates := "SrcType := Int" } EQ_Contact(in1 := "Valves Data".R9_XV02.STATUS, in2 := 1)
   END_RUNG wire#w6
   RUNG wire#w5
      { S7_Templates := "SrcType := Int" } EQ_Contact(in1 := "Valves Data".R9_XV03.STATUS, in2 := 1)
   END_RUNG wire#w6
   // the same network as SCL:
   IF "AlwaysTRUE" THEN
       #valve_R9_XV04("auto/manual" := "Valves Data"."A/M".R9,   // "valve"
                      open_auto := "R9_DATA".R9.UCHWS_CMD_2 OR "R9_DATA".R9.UCHWS_CMD_1,
                      open_man := "Valves Data".R9_XV04.MCMD AND NOT "dummy".R9.Intl_4,
                      fbk_open := "A/GLR_009_XV502_OFB",
                      fbk_close := "A/GLR_009_XV502_CFB",
                      reset := "Valves Data".R9_XV04.RESET OR "R9_DATA".R9.Reset,
                      intl := NOT "DI_INPUTS".R9_INPUTS_RUA.EMG_PB,
                      Mon_En := 1,
                      mon_sp := "Valves Data".R9_XV04.MON_TIME,
                      SEMI := "Valves Data".SEMI_AUTO.R9,
                      "open/close" => "A/GLR_009_XV502_CMD",
                      FAIL_TO_OPEN => "Valves Data".R9_VALVE_FAULT.XV04_FAIL_TO_OPEN,
                      FAIL_TO_CLOSE => "Valves Data".R9_VALVE_FAULT.XV04_FAIL_TO_CLOSE,
                      status => "Valves Data".R9_XV04.STATUS);
   END_IF;
   "dummy".R9.Intl_4 := "AlwaysTRUE" AND (("Valves Data".R9_XV01.STATUS = 1) OR ("Valves Data".R9_XV02.STATUS = 1) OR ("Valves Data".R9_XV03.STATUS = 1));
END_REGION

REGION Network 93: R9_XV05
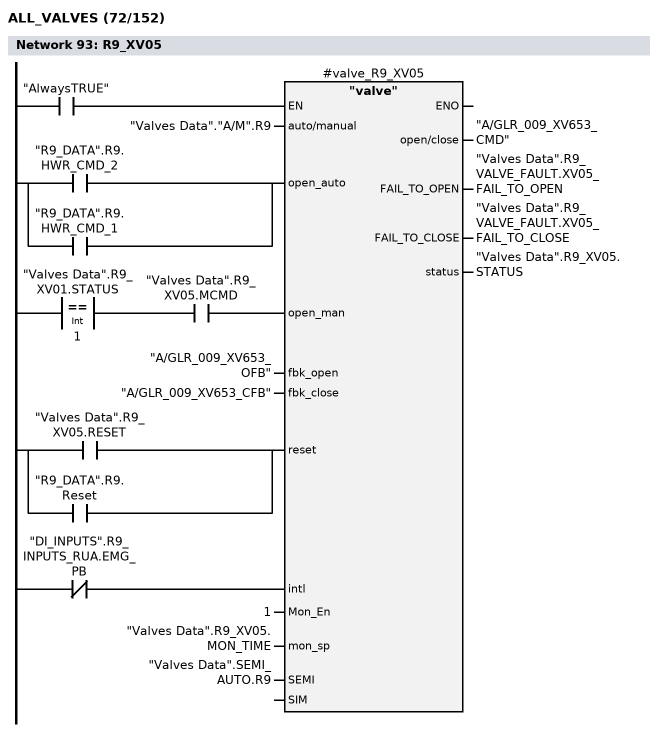
   RUNG wire#powerrail
      Contact( "AlwaysTRUE" )
      #valve_R9_XV05(open_auto := wire#w1, open_man := wire#w2, reset := wire#w3, intl := wire#w4, "auto/manual" := "Valves Data"."A/M".R9, fbk_open := "A/GLR_009_XV653_OFB", fbk_close := "A/GLR_009_XV653_CFB", Mon_En := 1, mon_sp := "Valves Data".R9_XV05.MON_TIME, SEMI := "Valves Data".SEMI_AUTO.R9, SIM :=, "open/close" => "A/GLR_009_XV653_CMD", FAIL_TO_OPEN => "Valves Data".R9_VALVE_FAULT.XV05_FAIL_TO_OPEN, FAIL_TO_CLOSE => "Valves Data".R9_VALVE_FAULT.XV05_FAIL_TO_CLOSE, status => "Valves Data".R9_XV05.STATUS)
   END_RUNG
   RUNG wire#powerrail
      Contact( "R9_DATA".R9.HWR_CMD_2 )
   END_RUNG wire#w1
   RUNG wire#powerrail
      Contact( "R9_DATA".R9.HWR_CMD_1 )
   END_RUNG wire#w1
   RUNG wire#powerrail
      { S7_Templates := "SrcType := Int" } EQ_Contact(in1 := "Valves Data".R9_XV01.STATUS, in2 := 1)
      Contact( "Valves Data".R9_XV05.MCMD )
   END_RUNG wire#w2
   RUNG wire#powerrail
      Contact( "Valves Data".R9_XV05.RESET )
   END_RUNG wire#w3
   RUNG wire#powerrail
      Contact( "R9_DATA".R9.Reset )
   END_RUNG wire#w3
   RUNG wire#powerrail
      I_Contact( "DI_INPUTS".R9_INPUTS_RUA.EMG_PB )
   END_RUNG wire#w4
   // the same network as SCL:
   IF "AlwaysTRUE" THEN
       #valve_R9_XV05("auto/manual" := "Valves Data"."A/M".R9,   // "valve"
                      open_auto := "R9_DATA".R9.HWR_CMD_2 OR "R9_DATA".R9.HWR_CMD_1,
                      open_man := ("Valves Data".R9_XV01.STATUS = 1) AND "Valves Data".R9_XV05.MCMD,
                      fbk_open := "A/GLR_009_XV653_OFB",
                      fbk_close := "A/GLR_009_XV653_CFB",
                      reset := "Valves Data".R9_XV05.RESET OR "R9_DATA".R9.Reset,
                      intl := NOT "DI_INPUTS".R9_INPUTS_RUA.EMG_PB,
                      Mon_En := 1,
                      mon_sp := "Valves Data".R9_XV05.MON_TIME,
                      SEMI := "Valves Data".SEMI_AUTO.R9,
                      "open/close" => "A/GLR_009_XV653_CMD",
                      FAIL_TO_OPEN => "Valves Data".R9_VALVE_FAULT.XV05_FAIL_TO_OPEN,
                      FAIL_TO_CLOSE => "Valves Data".R9_VALVE_FAULT.XV05_FAIL_TO_CLOSE,
                      status => "Valves Data".R9_XV05.STATUS);
   END_IF;
END_REGION

REGION Network 94: R9_XV06
